(* IEC 61131-3 sources: daoli-st-library/DL_Process (part 41) *)

(* ---- FB_DL_LyoShelfTempRampCtrl.st ---- *)
(*
  Name: FB_DL_LyoShelfTempRampCtrl
  Category: DL_Process
  Version: 1.0.0
  Round: R91 / 2026-11-25
  开源溯源：clean-room 自研（族 制药冻干真空冷冻干燥，ST 开源生态实测 0 命中，无外部代码引入）
  功能：1) 搁板温度斜坡发生器：设定值 fSetpointC 以 fRateUpKmin / fRateDownKmin 的斜率
           逐拍逼近目标温度 fTargetC，每拍增量 = 斜率[K/min] / 60 * fCycleS[s]，
           接近目标时按「不越过目标」截断，天然消除斜坡积分超调。
        2) 超调抑制：实测温度 fActualC 越过目标温度且超出 fOverShootLimitK 并持续 DL_OV_DELAY 后，
           判超调故障并锁码 —— 这是加热回路失控（固态继电器击穿或传感器脱落）的实证判据。
        3) 斜率上下限约束：fRateUpKmin / fRateDownKmin 必须落在 (0.0, DL_RATE_HI_KMIN] 内，
           越域判故障码（斜率为零会让设定值永不到达，斜率过大会撕裂制品冰晶结构）。
  边界条件：1) 非有限值闸：目标温度、实测温度、两路斜率、周期先过 NOT(x > -DL_BIG AND x < DL_BIG)，
           同时拦 NaN 与 Inf；命中即判故障码 0213 并进故障相，
           绝不把 NaN 写进设定值（NaN 一旦进入斜坡状态量会永久污染积分链，R19）。
        2) 周期入参闸（R21）：fCycleS <= 0.0 或非有限时改用缺省 DL_CYCLE_DEF = 0.1 s 并置信息级码 0212，
           不静默改用。
        3) 斜率零闸：两路斜率均须 > DL_EPS，否则判故障码 0214（斜坡永不推进 = 温度控制静默失效）。
        4) 超调判据去抖：超调为瞬时量，必须经 tonOver 去抖后才升级为故障，避免单点尖峰误停。
        5) 单点赋值（R26）：fSetpointC 只在段 7 统一出口写一次；内部设定量 _fSpC 才是逐拍累加的对象。
        6) 故障解除路径：故障相内 xReset 上升沿 AND NOT xFault AND 入参有限 → 清锁存回待机，
           回待机后设定值跟随实测温度重新起步（无扰切换），不从零开始。
        7) 状态机兜底：CASE 全态覆盖 + ELSE 强制回故障相并置码 0217、清全部输出。
  量纲自证：斜率 [K/min] / 60 [s/min] * fCycleS [s] = 每拍增量 [K]，
           与 fSetpointC / fTargetC / fOverShootLimitK 同量纲 [K]（degC 差值以 K 计），量纲合法。
  码表 Error codes（本件子带 0091_021x，故障级一律 3 行内置 _uFault/_bFault/_eState）:
    16#0091_0211 信息级：使能关闭，设定值冻结在当下（不置故障位）
    16#0091_0212 信息级：周期入参非法，已按缺省 0.1 s 折算（不置故障位）
    16#0091_0213 故障级：温度或斜率入参非有限（NaN / Inf）
    16#0091_0214 故障级：斜率组态越域（为零或超物理上限）
    16#0091_0215 故障级：实测温度超调越限（加热回路失控判据）
    16#0091_0216 故障级：外部故障输入 xFault
    16#0091_0217 故障级：状态机落 ELSE 兜底（非法相位 ID）

  修订历史 Revision :
    2026-11-25  v1.0.0  R91 首版
*)

TYPE E_DL_LyoShelfRampState :
(
    eLyoRampIdle  := 0,     // 待机：使能关闭，设定值冻结 / Idle, disabled and setpoint frozen
    eLyoRampHeat  := 10,    // 升温：设定值按升斜率逼近目标 / Heating, setpoint ramps up to target
    eLyoRampCool  := 20,    // 降温：设定值按降斜率逼近目标 / Cooling, setpoint ramps down to target
    eLyoRampHold  := 30,    // 保持：设定值已达目标，进入保温带 / Hold, setpoint on target within the band
    eLyoRampFault := 90     // 故障：锁存待解除 / Fault, latched awaiting release
);
END_TYPE

FUNCTION_BLOCK FB_DL_LyoShelfTempRampCtrl
VAR_INPUT
    xEnable        : BOOL;    // 斜坡控制使能 [bool] / Ramp control enable [bool]
    xReset         : BOOL;    // 故障复位（上升沿有效）[bool] / Fault reset, rising edge [bool]
    xFault         : BOOL;    // 外部故障汇总 [bool] / External fault aggregate [bool]
    fTargetC       : REAL;    // 搁板目标温度 [degC] / Shelf target temperature [degC]
    fActualC       : REAL;    // 搁板实测温度 [degC] / Shelf measured temperature [degC]
    fRateUpKmin    : REAL;    // 允许升温斜率 [K/min] / Permitted heating rate [K/min]
    fRateDownKmin  : REAL;    // 允许降温斜率 [K/min] / Permitted cooling rate [K/min]
    fCycleS        : REAL;    // 任务周期 [s] / Task cycle time [s]
    fBandK         : REAL;    // 到温判定带宽 [K] / At-target band width [K]
    fOverShootLimitK : REAL;  // 允许超调量 [K] / Permitted overshoot [K]
END_VAR
VAR_OUTPUT
    fSetpointC     : REAL;    // 搁板温度设定值 [degC] / Shelf temperature setpoint [degC]
    xHeating       : BOOL;    // 升温方向标志 [bool] / Heating direction flag [bool]
    xCooling       : BOOL;    // 降温方向标志 [bool] / Cooling direction flag [bool]
    xInBand        : BOOL;    // 已进入到温带 [bool] / Within the at-target band [bool]
    xOverShoot     : BOOL;    // 超调越限标志（已去抖）[bool] / Overshoot flag, debounced [bool]
    eState         : E_DL_LyoShelfRampState;   // 状态出口，段尾单点映射 / State outlet, single-point mapped
    nErrId         : UDINT;   // 事件码，0 = 无事件 / Event code, 0 = none
END_VAR
VAR
    tonOver        : TON;     // 超调去抖定时 [TIME] / Overshoot debounce timer
    rtReset        : R_TRIG;  // 复位上升沿检测 [bool] / Reset rising edge detector
    _eState        : E_DL_LyoShelfRampState := E_DL_LyoShelfRampState.eLyoRampIdle;   // 内部相位（CASE 唯一写入目标）
    _fSpC          : REAL := 0.0;   // 内部设定值状态量（逐拍累加对象）[degC] / Internal setpoint state [degC]
    _fStepK        : REAL := 0.0;   // 本拍温度增量 [K] / Temperature increment this cycle [K]
    _fCycleUseS    : REAL := 0.1;   // 实际使用的周期值 [s] / Cycle time actually used [s]
    _bFinOk        : BOOL := FALSE; // 实值入参有限性总闸结果 / Finiteness gate aggregate result
    _bRateOk       : BOOL := FALSE; // 斜率组态域闸结果 / Ramp rate domain gate result
    _bCycleBad     : BOOL := FALSE; // 周期入参非法标志 [bool] / Cycle input invalid flag [bool]
    _bOverRaw      : BOOL := FALSE; // 超调原始判据（未去抖）[bool] / Raw overshoot criterion
    _bFault        : BOOL := FALSE; // 故障锁存位 [bool] / Latched fault flag [bool]
    _bSpInit       : BOOL := FALSE; // 设定值已初始化标志 [bool] / Setpoint initialised flag [bool]
    _uInfo         : UDINT := 16#0000_0000;   // 信息码，每拍重算 / Info code, recomputed every cycle
    _uFault        : UDINT := 16#0000_0000;   // 故障码锁存 / Latched fault code
END_VAR
VAR CONSTANT
    DL_EPS         : REAL := 1.0E-9;      // 数值零闸阈值 [-] / Numeric zero gate threshold [-]
    DL_BIG         : REAL := 1.0E12;      // 非有限值闸量级上限 [-] / Finiteness gate magnitude [-]
    DL_CYCLE_DEF   : REAL := 0.1;         // 缺省任务周期 [s] / Default task cycle time [s]
    DL_CYCLE_MIN   : REAL := 0.001;       // 周期合理下限 [s] / Cycle time reasonable low bound [s]
    DL_CYCLE_MAX   : REAL := 10.0;        // 周期合理上限 [s] / Cycle time reasonable high bound [s]
    DL_SEC_PER_MIN : REAL := 60.0;        // 分钟到秒的时基折算 [s/min] / Seconds per minute [s/min]
    DL_RATE_HI_KMIN: REAL := 10.0;        // 允许斜率物理上限 [K/min] / Ramp rate physical upper bound [K/min]
    DL_OV_DELAY    : TIME := T#10S;       // 超调去抖窗 [TIME] / Overshoot debounce window [TIME]
    DL_T_SPAN      : REAL := 300.0;       // 温度量级闸跨度 [degC] / Temperature magnitude gate span [degC]
END_VAR

(* —— 段 0：单拍量预清零（锁存量 _uFault/_bFault/_bSpInit 不入清单，R187①） —— *)
_uInfo := 16#0000_0000;                     // 信息码每拍重算 / Info code recomputed
nErrId := 16#0000_0000;                     // 事件码缺省无事件 / Event code defaults to none

(* —— 段 1：周期入参闸（R21：非法周期不静默，改用缺省并置信息码） —— *)
_bCycleBad := NOT (fCycleS > -DL_BIG AND fCycleS < DL_BIG)
              OR (fCycleS < DL_CYCLE_MIN) OR (fCycleS > DL_CYCLE_MAX);
IF _bCycleBad THEN
    _fCycleUseS := DL_CYCLE_DEF;            // 非法周期一律用缺省 0.1 s
    _uInfo := 16#0091_0212;                 // 信息级：周期入参非法，已用缺省（不置故障位）
ELSE
    _fCycleUseS := fCycleS;                 // 合法周期原值使用
END_IF

(* —— 段 2：非有限值闸与斜率域闸（R19：不把 NaN 写进斜坡状态量） —— *)
_bFinOk := (fTargetC > -DL_BIG) AND (fTargetC < DL_BIG)
           AND (fActualC > -DL_BIG) AND (fActualC < DL_BIG)
           AND (fRateUpKmin > -DL_BIG) AND (fRateUpKmin < DL_BIG)
           AND (fRateDownKmin > -DL_BIG) AND (fRateDownKmin < DL_BIG)
           AND (fBandK > -DL_BIG) AND (fBandK < DL_BIG)
           AND (fOverShootLimitK > -DL_BIG) AND (fOverShootLimitK < DL_BIG);
_bRateOk := (fRateUpKmin > DL_EPS) AND (fRateUpKmin <= DL_RATE_HI_KMIN)
            AND (fRateDownKmin > DL_EPS) AND (fRateDownKmin <= DL_RATE_HI_KMIN)
            AND (fBandK > DL_EPS) AND (fOverShootLimitK > DL_EPS)
            AND (ABS(fTargetC) <= DL_T_SPAN) AND (ABS(fActualC) <= DL_T_SPAN);

(* —— 段 3：超调原始判据（仅升温方向有意义：实测高于目标且超出允许量） —— *)
_bOverRaw := _bFinOk AND _bRateOk
             AND ((fActualC - fTargetC) > fOverShootLimitK);

(* —— 段 4：边沿与定时器无条件周期刷新（R7：调用语句不得置于 IF/CASE 内） —— *)
rtReset(CLK := xReset);                                             // 复位上升沿，每拍必调
tonOver(IN := _bOverRaw AND (NOT _bFault), PT := DL_OV_DELAY);      // 超调去抖

(* —— 段 5：全局故障拦截（优先级最高；已锁存则不再改写码值，禁同拍抹除） —— *)
IF xFault AND (NOT _bFault) THEN
    _uFault := 16#0091_0216;                // 故障级：外部故障输入
    _bFault := TRUE;                        // 锁存（3 行内置，R45 配对）
    _eState := E_DL_LyoShelfRampState.eLyoRampFault;
END_IF
IF (NOT _bFinOk) AND (NOT _bFault) THEN
    _uFault := 16#0091_0213;                // 故障级：入参非有限（独立成因，R190）
    _bFault := TRUE;                        // 锁存
    _eState := E_DL_LyoShelfRampState.eLyoRampFault;
END_IF
IF (NOT _bRateOk) AND _bFinOk AND (NOT _bFault) THEN
    _uFault := 16#0091_0214;                // 故障级：斜率组态越域（独立成因，R190）
    _bFault := TRUE;                        // 锁存
    _eState := E_DL_LyoShelfRampState.eLyoRampFault;
END_IF
IF tonOver.Q AND (NOT _bFault) THEN
    _uFault := 16#0091_0215;                // 故障级：实测温度超调越限
    _bFault := TRUE;                        // 锁存
    _eState := E_DL_LyoShelfRampState.eLyoRampFault;
END_IF

(* —— 段 6：设定值起步（首次使能或无扰复位时以实测温度初始化，避免设定值从零跳变） —— *)
IF (NOT _bSpInit) AND _bFinOk THEN
    _fSpC := fActualC;                      // 无扰起步：设定值跟随实测温度
    _bSpInit := TRUE;                       // 标记已初始化
END_IF

(* —— 段 7：相位机（只做迁移与内部设定值更新；出口在段 9 单点映射） —— *)
CASE _eState OF

E_DL_LyoShelfRampState.eLyoRampIdle:
    IF NOT xEnable THEN
        _uInfo := 16#0091_0211;             // 信息级：使能关闭，设定值冻结（不置故障位）
    ELSIF (fTargetC - _fSpC) > fBandK THEN
        _eState := E_DL_LyoShelfRampState.eLyoRampHeat;       // 目标高于设定值：进升温相
    ELSIF (_fSpC - fTargetC) > fBandK THEN
        _eState := E_DL_LyoShelfRampState.eLyoRampCool;       // 目标低于设定值：进降温相
    ELSE
        _eState := E_DL_LyoShelfRampState.eLyoRampHold;       // 已在带内：进保持相
    END_IF

E_DL_LyoShelfRampState.eLyoRampHeat:
    IF (NOT xEnable) OR _bFault THEN
        _uInfo := 16#0091_0211;             // 信息级：失能即冻结设定值
        _eState := E_DL_LyoShelfRampState.eLyoRampIdle;
    ELSE
        _fStepK := fRateUpKmin / DL_SEC_PER_MIN * _fCycleUseS;                 // 每拍升温增量 [K]
        _fSpC := _fSpC + _fStepK;                                             // 累加
        IF _fSpC >= fTargetC THEN
            _fSpC := fTargetC;              // 不越过目标：天然消除斜坡超调
            _eState := E_DL_LyoShelfRampState.eLyoRampHold;
        END_IF
    END_IF

E_DL_LyoShelfRampState.eLyoRampCool:
    IF (NOT xEnable) OR _bFault THEN
        _uInfo := 16#0091_0211;             // 信息级：失能即冻结设定值
        _eState := E_DL_LyoShelfRampState.eLyoRampIdle;
    ELSE
        _fStepK := fRateDownKmin / DL_SEC_PER_MIN * _fCycleUseS;               // 每拍降温增量 [K]
        _fSpC := _fSpC - _fStepK;                                             // 累减
        IF _fSpC <= fTargetC THEN
            _fSpC := fTargetC;              // 不越过目标：天然消除斜坡超调
            _eState := E_DL_LyoShelfRampState.eLyoRampHold;
        END_IF
    END_IF

E_DL_LyoShelfRampState.eLyoRampHold:
    IF (NOT xEnable) OR _bFault THEN
        _uInfo := 16#0091_0211;             // 信息级：失能即回待机
        _eState := E_DL_LyoShelfRampState.eLyoRampIdle;
    ELSIF (fTargetC - _fSpC) > fBandK THEN
        _eState := E_DL_LyoShelfRampState.eLyoRampHeat;       // 目标抬高：重返升温相（判据在钉住之前取）
    ELSIF (_fSpC - fTargetC) > fBandK THEN
        _eState := E_DL_LyoShelfRampState.eLyoRampCool;       // 目标压低：重返降温相（判据在钉住之前取）
    ELSE
        _fSpC := fTargetC;                  // 带内才钉住设定值（避免判据恒真）
    END_IF

E_DL_LyoShelfRampState.eLyoRampFault:
    IF rtReset.Q AND (NOT xFault) AND _bFinOk AND _bRateOk THEN
        _bFault := FALSE;                   // 解除路径：复位沿 + 外部故障消失 + 入参与组态合法（可达，R188）
        _uFault := 16#0000_0000;            // 清锁存码
        _bSpInit := FALSE;                  // 强制无扰重启：设定值重新跟随实测温度
        _eState := E_DL_LyoShelfRampState.eLyoRampIdle;       // 回待机
    END_IF

ELSE
    _uFault := 16#0091_0217;                // 故障级：非法相位 ID 兜底
    _bFault := TRUE;                        // 锁存
    _eState := E_DL_LyoShelfRampState.eLyoRampFault;          // 强制回故障相

END_CASE

(* —— 段 8：后置段（设定值域兜底：非有限或越量级一律回落到实测温度） —— *)
IF NOT (_fSpC > -DL_BIG AND _fSpC < DL_BIG) THEN
    _fSpC := fActualC;                      // 内部状态自检：非有限即回落实测值
END_IF
(* —— 段 8.5：出口值域二阶终闸（R19 二阶形态）——
   一次闸的回退源是 fActualC，而 fActualC 本身也可能是非有限值（入参 NaN/Inf），
   回退后仍为 NaN，且 ABS(NaN) > DL_T_SPAN 恒假会绕过越量级钳制，NaN 直穿设定值出口。
   故必须对「回退之后」的值再做一次判据与钳制，才真正闸断实值通路。 *)
IF NOT (_fSpC >= -DL_T_SPAN AND _fSpC <= DL_T_SPAN) THEN
    _fSpC := 0.0;                           // 双源皆非有限：0 degC 安全位 / Both sources non-finite: 0 degC safe
END_IF
IF ABS(_fSpC) > DL_T_SPAN THEN
    _fSpC := LIMIT(-DL_T_SPAN, _fSpC, DL_T_SPAN);   // 越量级钳制，防积分链发散
END_IF

(* —— 段 9：出口单点映射（名实同源；方向位由设定值与目标差导出，故障侧全清） —— *)
IF _bFault THEN
    IF (fActualC >= -DL_T_SPAN) AND (fActualC <= DL_T_SPAN) THEN
        fSetpointC := fActualC;             // 故障侧优先回落实测温度（有限时保持原语义：冻结在实测）
    ELSE
        fSetpointC := _fSpC;                // 实测非有限时回落到已过二阶终闸的安全值，绝不输出 NaN
    END_IF;
    xHeating := FALSE;                      // 故障侧方向位清零
    xCooling := FALSE;                      // 故障侧方向位清零
    xInBand := FALSE;                       // 故障侧到温位清零
ELSE
    fSetpointC := _fSpC;                    // 正常侧设定值出口
    xHeating := (_eState = E_DL_LyoShelfRampState.eLyoRampHeat);      // 升温方向位
    xCooling := (_eState = E_DL_LyoShelfRampState.eLyoRampCool);      // 降温方向位
    xInBand := (_eState = E_DL_LyoShelfRampState.eLyoRampHold)        // 到温带：保持相且实测在带内
               AND (ABS(fActualC - fTargetC) <= fBandK);
END_IF
xOverShoot := tonOver.Q;                    // 超调位出口（已去抖）
eState := _eState;                          // 状态出口单点映射
IF _bFault THEN
    nErrId := _uFault;                      // 故障锁存码回放（不在故障相按当下输入重推断）
ELSE
    nErrId := _uInfo;                       // 信息码
END_IF

END_FUNCTION_BLOCK

(* ---- FB_DL_LyoVacuumPullSeq.st ---- *)
(*
  Name: FB_DL_LyoVacuumPullSeq
  Category: DL_Process
  Version: 1.0.0
  Round: R91 / 2026-11-25
  开源溯源：clean-room 自研（族 制药冻干真空冷冻干燥，ST 开源生态实测 0 命中，无外部代码引入）
  功能：1) 抽真空状态机，六相推进：待机 → 粗抽 → 精抽 → 保持 → 就绪 → （通气）。
           待机相等 xStart 上升沿；腔体压力已低于粗抽目标时跳过粗抽相（信息级码 0231 声明跳过）；
           粗抽相开粗抽泵阀组，压力降到 fRoughTargetMbar 即转精抽；精抽相关粗抽阀、开精抽阀，
           压力降到 fFineTargetMbar 即转保持相；保持相关全部抽气、观察 tHoldS 内压力升幅，
           升幅 <= fHoldRiseMaxMbar 判真空保持合格，置 xHoldOk 并进就绪相；
           就绪相保持 xReady 直到 xStart 撤下；撤令后进通气相复压并回待机。
        2) 泵故障兜底：粗抽/精抽/保持三相内，泵运行反馈丢失或泵过载上升即锁码 0237 并立即进故障相，
           同时撤销全部抽气命令、不打开通气阀（避免带故障强行复压把油雾带入腔体）。
        3) 每相独立超时 + 整序总超时：四个相定时器各配一个「定时 + 裕量」超时点，
           tonTotal 兜底整序总时长；保持相另配真空上升超限判据（0234）与稳定超时（0235）双归因。
  边界条件：1) 非有限值闸：压力、三个目标限值先过 NOT(x > -DL_BIG AND x < DL_BIG)，同时拦 NaN 与 Inf；
           命中即锁码 0239 进故障相，绝不把 NaN 拿去与真空目标比较（NaN 比较恒假会让抽气永不停止，R19）。
        2) 组态域闸：三个压力阈须满足 0.0 < fFineTargetMbar < fRoughTargetMbar（真空度方向由粗到精），
           fHoldRiseMaxMbar > DL_EPS，越域锁码 0239（组态错误与入参非有限共用同一归因码前缀，
           但内部用两个独立成员区分，见 _bCfgOk / _bFinOk）。
        3) 压力单调性：抽气相内压力不得上升；若在粗抽/精抽相检测到压力高于本相入口压力且超过
           DL_PRESS_TOL，视为泵失效实测证据，锁码 0232 / 0233（与超时归因区分：这里不是等不到，而是反向）。
        4) 时间参数零闸：tRoughS / tFineS / tHoldS <= T#0S 时对应相定时器立即置 Q（等价跳过），
           属调试合法组态；但保持相零窗会使升幅判据恒成立，故保持相入口对 tHoldS 做显式零闸 → 锁码 0235。
        5) 定时器周期刷新（R7）：八个 TON 与复位边沿全部在 CASE 之外无条件调用。
        6) 故障解除路径：故障相内 xReset 上升沿 AND NOT xFault AND 入参/组态合法 → 清锁存回待机，
           回待机后必须重新给 xStart 上升沿才能再启动（不自恢复）。
        7) 状态机兜底：CASE 全态覆盖 + ELSE 强制回故障相并置码 0240、清全部输出。
        8) 输出安全初值（R25）：三个阀门命令初值 FALSE、xReady 初值 FALSE，待机相显式赋值。
  量纲自证：fChamberPressMbar / fRoughTargetMbar / fFineTargetMbar / fHoldRiseMaxMbar 全为压力 [mbar]，
           比较两侧同量纲；升幅 = 保持末压力 − 保持初压力，仍为 [mbar]；
           所有时间引脚为 [TIME]，相超时点 = [TIME] + [TIME] = [TIME]，与 TON 的 PT 同量纲。
  码表 Error codes（本件子带 0091_024x，故障级一律 3 行内置 _uFault/_bFault/_eState）:
    16#0091_0231 信息级：腔体压力已低于粗抽目标，跳过粗抽相（不置故障位）
    16#0091_0232 故障级：粗抽相超时（定时到但未达粗抽目标）
    16#0091_0233 故障级：精抽相超时（定时到但未达精抽目标）
    16#0091_0234 故障级：保持相真空度上升超限（泄漏或放气）
    16#0091_0235 故障级：保持相超时或保持窗为零（压力未稳定/判据恒真）
    16#0091_0236 故障级：整序总超时
    16#0091_0237 故障级：泵运行反馈丢失或泵过载
    16#0091_0238 故障级：外部故障输入 xFault
    16#0091_0239 故障级：压力/限值入参非有限，或压力阈组态越域
    16#0091_0240 故障级：状态机落 ELSE 兜底（非法相位 ID）
    16#0091_0241 信息级：就绪保持中，等待撤令（不置故障位）
    16#0091_0242 信息级：通气复压相进行中（不置故障位）
    16#0091_0243 信息级：泵未就绪（无运行反馈或过载），暂不启动抽气（不置故障位）
    16#0091_0244 故障级：粗抽相压力反向上升（泵失效实证，与超时成因分离）
    16#0091_0245 故障级：精抽相压力反向上升（泄漏或阀未开，与超时成因分离）
    16#0091_0246 故障级：通气相超时（复压未完成）

  修订历史 Revision :
    2026-11-25  v1.0.0  R91 首版
*)

TYPE E_DL_LyoVacuumPullState :
(
    eLyoVacIdle  := 0,      // 待机：等启动上升沿 / Idle, awaiting the start rising edge
    eLyoVacRough := 10,     // 粗抽：粗抽泵组开，降到粗抽目标 / Rough pull, pump group on
    eLyoVacFine  := 20,     // 精抽：关粗抽阀开精抽阀，降到精抽目标 / Fine pull, fine valve open
    eLyoVacHold  := 30,     // 保持：关全部抽气，测压力升幅 / Hold, all pumping off, rise measured
    eLyoVacReady := 40,     // 就绪：真空保持合格，保持到位 / Ready, vacuum hold accepted
    eLyoVacVent  := 50,     // 通气：开通气阀复压回待机 / Vent, repressurising back to idle
    eLyoVacFault := 90      // 故障：锁存待解除 / Fault, latched awaiting release
);
END_TYPE

FUNCTION_BLOCK FB_DL_LyoVacuumPullSeq
VAR_INPUT
    xStart           : BOOL;   // 抽真空启动指令（上升沿有效）[bool] / Vacuum pull start, edge triggered [bool]
    xReset           : BOOL;   // 故障复位（上升沿有效）[bool] / Fault reset, rising edge [bool]
    xFault           : BOOL;   // 外部故障汇总 [bool] / External fault aggregate [bool]
    xPumpRunFb       : BOOL;   // 真空泵运行反馈 [bool] / Vacuum pump running feedback [bool]
    xPumpOverload    : BOOL;   // 真空泵过载信号 [bool] / Vacuum pump overload signal [bool]
    fChamberPressMbar : REAL;  // 腔体实测压力 [mbar] / Measured chamber pressure [mbar]
    fRoughTargetMbar : REAL;   // 粗抽目标压力 [mbar] / Rough pull target pressure [mbar]
    fFineTargetMbar  : REAL;   // 精抽目标压力 [mbar] / Fine pull target pressure [mbar]
    fHoldRiseMaxMbar : REAL;   // 保持相允许压力升幅 [mbar] / Permitted pressure rise during hold [mbar]
    tRoughS          : TIME;   // 粗抽相设定时长 [TIME] / Rough pull phase duration [TIME]
    tFineS           : TIME;   // 精抽相设定时长 [TIME] / Fine pull phase duration [TIME]
    tHoldS           : TIME;   // 保持相设定时长 [TIME] / Hold phase duration [TIME]
END_VAR
VAR_OUTPUT
    xRoughValveCmd   : BOOL;   // 粗抽阀命令（安全侧：故障时关）[bool] / Rough valve command, fail-safe [bool]
    xFineValveCmd    : BOOL;   // 精抽阀命令（安全侧：故障时关）[bool] / Fine valve command, fail-safe [bool]
    xVentValveCmd    : BOOL;   // 通气阀命令（安全侧：故障时关）[bool] / Vent valve command, fail-safe [bool]
    xHoldOk          : BOOL;   // 真空保持判据通过（跨相保持）[bool] / Vacuum hold accepted, held across phases [bool]
    xReady           : BOOL;   // 抽真空就绪保持位 [bool] / Vacuum ready held flag [bool]
    xBusy            : BOOL;   // 抽真空进行中 [bool] / Vacuum pull busy [bool]
    eState           : E_DL_LyoVacuumPullState;   // 状态出口，段尾单点映射 / State outlet, single-point mapped
    nErrId           : UDINT;  // 事件码，0 = 无事件 / Event code, 0 = none
END_VAR
VAR
    tonRough         : TON;    // 粗抽相正常定时 [TIME] / Rough pull phase timer
    tonRoughOv       : TON;    // 粗抽相超时定时 [TIME] / Rough pull phase overrun timer
    tonFine          : TON;    // 精抽相正常定时 [TIME] / Fine pull phase timer
    tonFineOv        : TON;    // 精抽相超时定时 [TIME] / Fine pull phase overrun timer
    tonHold          : TON;    // 保持相正常定时 [TIME] / Hold phase timer
    tonHoldOv        : TON;    // 保持相超时定时 [TIME] / Hold phase overrun timer
    tonVent          : TON;    // 通气相正常定时 [TIME] / Vent phase timer
    tonVentOv        : TON;    // 通气相超时定时 [TIME] / Vent phase overrun timer
    tonTotal         : TON;    // 整序总超时定时 [TIME] / Whole-sequence total timeout timer
    rtStart          : R_TRIG; // 启动上升沿检测 [bool] / Start rising edge detector
    rtReset          : R_TRIG; // 复位上升沿检测 [bool] / Reset rising edge detector
    _eState          : E_DL_LyoVacuumPullState := E_DL_LyoVacuumPullState.eLyoVacIdle;   // 内部相位（CASE 唯一写入目标）
    _fPressEntryMbar : REAL := 0.0;   // 本相入口压力快照 [mbar] / Pressure snapshot at phase entry [mbar]
    _fHoldStartMbar  : REAL := 0.0;   // 保持相起点压力快照 [mbar] / Pressure snapshot at hold start [mbar]
    _fRiseMbar       : REAL := 0.0;   // 保持相压力升幅 [mbar] / Pressure rise during the hold phase [mbar]
    _bFinOk          : BOOL := FALSE; // 实值入参有限性总闸结果 / Finiteness gate aggregate result
    _bCfgOk          : BOOL := FALSE; // 压力阈组态域闸结果 / Pressure threshold domain gate result
    _bPumpOk         : BOOL := FALSE; // 泵健康（运行反馈有且无过载）[bool] / Pump healthy flag [bool]
    _bActive         : BOOL := FALSE; // 序激活（粗抽至通气五相之一）[bool] / Sequence active flag [bool]
    _bHoldL          : BOOL := FALSE; // 保持合格位锁存（跨相保持）[bool] / Hold-accepted latch [bool]
    _bFault          : BOOL := FALSE; // 故障锁存位 [bool] / Latched fault flag [bool]
    _uInfo           : UDINT := 16#0000_0000;   // 信息码，每拍重算 / Info code, recomputed every cycle
    _uFault          : UDINT := 16#0000_0000;   // 故障码锁存 / Latched fault code
END_VAR
VAR CONSTANT
    DL_EPS         : REAL := 1.0E-9;      // 数值零闸阈值 [-] / Numeric zero gate threshold [-]
    DL_BIG         : REAL := 1.0E12;      // 非有限值闸量级上限 [-] / Finiteness gate magnitude [-]
    DL_PRESS_TOL   : REAL := 0.05;        // 抽气相压力反向容差 [mbar] / Reverse-trend tolerance while pumping [mbar]
    DL_P_HI        : REAL := 1100.0;      // 压力量级闸上限（略高于常压）[mbar] / Pressure magnitude gate upper bound [mbar]
    DL_OVER_MARGIN : TIME := T#60S;       // 相超时相对正常定时的裕量 [TIME] / Phase overrun margin [TIME]
    DL_TOTAL_MAX   : TIME := T#4H;        // 整序总超时上限 [TIME] / Whole-sequence total timeout [TIME]
    DL_ZERO_PRES   : REAL := 0.0;         // 压力零基准 [mbar] / Zero pressure reference [mbar]
END_VAR

(* —— 段 0：单拍量预清零（锁存量 _uFault/_bFault/_bHoldL 不入清单，R187①） —— *)
_uInfo := 16#0000_0000;                     // 信息码每拍重算 / Info code recomputed
nErrId := 16#0000_0000;                     // 事件码缺省无事件 / Event code defaults to none

(* —— 段 1：非有限值闸与组态域闸（R19：不拿 NaN 去比较真空目标） —— *)
_bFinOk := (fChamberPressMbar > -DL_BIG) AND (fChamberPressMbar < DL_BIG)
           AND (fRoughTargetMbar > -DL_BIG) AND (fRoughTargetMbar < DL_BIG)
           AND (fFineTargetMbar > -DL_BIG) AND (fFineTargetMbar < DL_BIG)
           AND (fHoldRiseMaxMbar > -DL_BIG) AND (fHoldRiseMaxMbar < DL_BIG);
_bCfgOk := (fFineTargetMbar > DL_EPS)                       // 精抽目标须为正压
           AND (fFineTargetMbar < fRoughTargetMbar)         // 精抽必须比粗抽更深（方向由粗到精）
           AND (fRoughTargetMbar < DL_P_HI)                 // 粗抽目标须在压力量级内
           AND (fHoldRiseMaxMbar > DL_EPS);                 // 允许升幅须组态为正

(* —— 段 2：泵健康判据（运行反馈 + 过载；过载优先） —— *)
_bPumpOk := xPumpRunFb AND (NOT xPumpOverload);

(* —— 段 3：派生态（序激活、保持升幅） —— *)
_bActive := (_eState = E_DL_LyoVacuumPullState.eLyoVacRough)
            OR (_eState = E_DL_LyoVacuumPullState.eLyoVacFine)
            OR (_eState = E_DL_LyoVacuumPullState.eLyoVacHold)
            OR (_eState = E_DL_LyoVacuumPullState.eLyoVacReady)
            OR (_eState = E_DL_LyoVacuumPullState.eLyoVacVent);
_fRiseMbar := fChamberPressMbar - _fHoldStartMbar;          // 保持相压力升幅 [mbar]

(* —— 段 4：定时器与边沿无条件周期刷新（R7：调用语句不得置于 IF/CASE 内） —— *)
rtStart(CLK := xStart);                                                                   // 启动上升沿，每拍必调
rtReset(CLK := xReset);                                                                   // 复位上升沿，每拍必调
tonRough(IN := (_eState = E_DL_LyoVacuumPullState.eLyoVacRough), PT := tRoughS);          // 粗抽相正常定时
tonRoughOv(IN := (_eState = E_DL_LyoVacuumPullState.eLyoVacRough),
           PT := tRoughS + DL_OVER_MARGIN);                                               // 粗抽相超时点
tonFine(IN := (_eState = E_DL_LyoVacuumPullState.eLyoVacFine), PT := tFineS);             // 精抽相正常定时
tonFineOv(IN := (_eState = E_DL_LyoVacuumPullState.eLyoVacFine),
          PT := tFineS + DL_OVER_MARGIN);                                                 // 精抽相超时点
tonHold(IN := (_eState = E_DL_LyoVacuumPullState.eLyoVacHold), PT := tHoldS);             // 保持相正常定时
tonHoldOv(IN := (_eState = E_DL_LyoVacuumPullState.eLyoVacHold),
          PT := tHoldS + DL_OVER_MARGIN);                                                 // 保持相超时点
tonVent(IN := (_eState = E_DL_LyoVacuumPullState.eLyoVacVent), PT := tRoughS);            // 通气相正常定时（借用粗抽时长作复压窗）
tonVentOv(IN := (_eState = E_DL_LyoVacuumPullState.eLyoVacVent),
          PT := tRoughS + DL_OVER_MARGIN);                                                // 通气相超时点
tonTotal(IN := _bActive, PT := DL_TOTAL_MAX);                                             // 整序总超时

(* —— 段 5：全局故障拦截（优先级最高；已锁存则不再改写码值，禁同拍抹除） —— *)
IF xFault AND (NOT _bFault) THEN
    _uFault := 16#0091_0238;                // 故障级：外部故障输入
    _bFault := TRUE;                        // 锁存（3 行内置，R45 配对）
    _eState := E_DL_LyoVacuumPullState.eLyoVacFault;
END_IF
IF ((NOT _bFinOk) OR (NOT _bCfgOk)) AND (NOT _bFault) THEN
    _uFault := 16#0091_0239;                // 故障级：入参非有限或压力阈组态越域（同一码，成员已分离）
    _bFault := TRUE;                        // 锁存
    _eState := E_DL_LyoVacuumPullState.eLyoVacFault;
END_IF
IF tonTotal.Q AND _bActive AND (NOT _bFault) THEN
    _uFault := 16#0091_0236;                // 故障级：整序总超时
    _bFault := TRUE;                        // 锁存
    _eState := E_DL_LyoVacuumPullState.eLyoVacFault;
END_IF
IF (NOT _bPumpOk) AND _bActive AND (NOT _bFault)
   AND (_eState <> E_DL_LyoVacuumPullState.eLyoVacVent) THEN
    _uFault := 16#0091_0237;                // 故障级：泵反馈丢失或过载（通气相不需泵，故排除）
    _bFault := TRUE;                        // 锁存
    _eState := E_DL_LyoVacuumPullState.eLyoVacFault;
END_IF

(* —— 段 6：相位机（只做迁移与锁存；出口在段 8 单点映射） —— *)
CASE _eState OF

E_DL_LyoVacuumPullState.eLyoVacIdle:
    IF NOT xStart THEN
        _bHoldL := FALSE;                   // 撤令即清保持合格位，为下次抽真空重新武装
        _fPressEntryMbar := fChamberPressMbar;   // 待机相刷新入口压力快照（有限性由段 5 保证）
    ELSIF rtStart.Q AND _bFinOk AND _bCfgOk THEN
        _bHoldL := FALSE;                   // 新序开始：清保持合格位
        _fPressEntryMbar := fChamberPressMbar;   // 捕获入口压力，供粗抽反向判据使用
        IF fChamberPressMbar <= fRoughTargetMbar THEN
            _uInfo := 16#0091_0231;         // 信息级：已低于粗抽目标，声明跳过粗抽相
            _eState := E_DL_LyoVacuumPullState.eLyoVacFine;      // 直接进精抽相
        ELSE
            _eState := E_DL_LyoVacuumPullState.eLyoVacRough;     // 进粗抽相
        END_IF
    ELSIF NOT _bPumpOk THEN
        _uInfo := 16#0091_0243;             // 信息级：泵未就绪，暂不启动（不置故障位）
    END_IF

E_DL_LyoVacuumPullState.eLyoVacRough:
    IF tonRoughOv.Q THEN
        _uFault := 16#0091_0232;            // 故障级：粗抽相超时
        _bFault := TRUE;                    // 锁存
        _eState := E_DL_LyoVacuumPullState.eLyoVacFault;
    ELSIF (fChamberPressMbar - _fPressEntryMbar) > DL_PRESS_TOL THEN
        _uFault := 16#0091_0244;            // 故障级：粗抽中压力反向上升（泵失效实证，独立成因）
        _bFault := TRUE;                    // 锁存
        _eState := E_DL_LyoVacuumPullState.eLyoVacFault;
    ELSIF fChamberPressMbar <= fRoughTargetMbar THEN
        _fPressEntryMbar := fChamberPressMbar;                   // 达粗抽目标：刷新入口快照（迁移前一次性）
        _eState := E_DL_LyoVacuumPullState.eLyoVacFine;          // 进精抽相
    END_IF

E_DL_LyoVacuumPullState.eLyoVacFine:
    IF tonFineOv.Q THEN
        _uFault := 16#0091_0233;            // 故障级：精抽相超时
        _bFault := TRUE;                    // 锁存
        _eState := E_DL_LyoVacuumPullState.eLyoVacFault;
    ELSIF (fChamberPressMbar - _fPressEntryMbar) > DL_PRESS_TOL THEN
        _uFault := 16#0091_0245;            // 故障级：精抽中压力反向上升（泄漏或阀未开，独立成因）
        _bFault := TRUE;                    // 锁存
        _eState := E_DL_LyoVacuumPullState.eLyoVacFault;
    ELSIF fChamberPressMbar <= fFineTargetMbar THEN
        _fHoldStartMbar := fChamberPressMbar;                    // 达精抽目标：捕获保持相起点压力
        _eState := E_DL_LyoVacuumPullState.eLyoVacHold;          // 进保持相
    END_IF

E_DL_LyoVacuumPullState.eLyoVacHold:
    IF tHoldS <= T#0S THEN
        _uFault := 16#0091_0235;            // 故障级：保持窗为零，升幅判据恒成立（不可接受组态）
        _bFault := TRUE;                    // 锁存
        _eState := E_DL_LyoVacuumPullState.eLyoVacFault;
    ELSIF tonHoldOv.Q THEN
        _uFault := 16#0091_0235;            // 故障级：保持相超时（压力未稳定）
        _bFault := TRUE;                    // 锁存
        _eState := E_DL_LyoVacuumPullState.eLyoVacFault;
    ELSIF tonHold.Q THEN
        IF _fRiseMbar > fHoldRiseMaxMbar THEN
            _uFault := 16#0091_0234;        // 故障级：保持相真空度上升超限（泄漏/放气）
            _bFault := TRUE;                // 锁存
            _eState := E_DL_LyoVacuumPullState.eLyoVacFault;
        ELSE
            _bHoldL := TRUE;                // 真空保持合格：锁存（跨相保持）
            _eState := E_DL_LyoVacuumPullState.eLyoVacReady;     // 进就绪相
        END_IF
    END_IF

E_DL_LyoVacuumPullState.eLyoVacReady:
    IF NOT xStart THEN
        _bHoldL := FALSE;                   // 撤令：清保持合格位并进通气相
        _eState := E_DL_LyoVacuumPullState.eLyoVacVent;
    ELSE
        _uInfo := 16#0091_0241;             // 信息级：就绪保持中，等撤令（不置故障位）
    END_IF

E_DL_LyoVacuumPullState.eLyoVacVent:
    IF tonVentOv.Q THEN
        _uFault := 16#0091_0246;            // 故障级：通气相超时（复压未完成，独立成因）
        _bFault := TRUE;                    // 锁存
        _eState := E_DL_LyoVacuumPullState.eLyoVacFault;
    ELSIF tonVent.Q THEN
        _eState := E_DL_LyoVacuumPullState.eLyoVacIdle;          // 复压完成：回待机
    ELSE
        _uInfo := 16#0091_0242;             // 信息级：通气复压进行中（不置故障位）
    END_IF

E_DL_LyoVacuumPullState.eLyoVacFault:
    IF rtReset.Q AND (NOT xFault) AND _bFinOk AND _bCfgOk THEN
        _bFault := FALSE;                   // 解除路径：复位沿 + 外部故障消失 + 入参/组态合法（可达，R188）
        _uFault := 16#0000_0000;            // 清锁存码
        _bHoldL := FALSE;                   // 保持合格位一并清，避免故障后误报就绪
        _eState := E_DL_LyoVacuumPullState.eLyoVacIdle;          // 回待机，需新上升沿才可再启动
    END_IF

ELSE
    _uFault := 16#0091_0240;                // 故障级：非法相位 ID 兜底
    _bFault := TRUE;                        // 锁存
    _eState := E_DL_LyoVacuumPullState.eLyoVacFault;             // 强制回故障相

END_CASE

(* —— 段 7：后置段（压力快照域兜底：非有限即清零，防污染下拍反向判据） —— *)
IF NOT (_fPressEntryMbar > -DL_BIG AND _fPressEntryMbar < DL_BIG) THEN
    _fPressEntryMbar := DL_ZERO_PRES;       // 内部状态自检：非有限即清零
END_IF
IF NOT (_fHoldStartMbar > -DL_BIG AND _fHoldStartMbar < DL_BIG) THEN
    _fHoldStartMbar := DL_ZERO_PRES;        // 内部状态自检：非有限即清零
END_IF

(* —— 段 8：出口单点映射（名实同源；阀门由状态导出，故障侧一律关阀） —— *)
xRoughValveCmd := (_eState = E_DL_LyoVacuumPullState.eLyoVacRough) AND (NOT _bFault);    // 粗抽阀：仅粗抽相
xFineValveCmd := (_eState = E_DL_LyoVacuumPullState.eLyoVacFine) AND (NOT _bFault);      // 精抽阀：仅精抽相
xVentValveCmd := (_eState = E_DL_LyoVacuumPullState.eLyoVacVent) AND (NOT _bFault);      // 通气阀：仅通气相
xHoldOk := _bHoldL AND (NOT _bFault);                                                    // 保持合格位出口
xReady := (_eState = E_DL_LyoVacuumPullState.eLyoVacReady) AND _bHoldL AND (NOT _bFault);   // 就绪位出口
xBusy := _bActive AND (NOT _bFault);                                                     // 进行中出口
eState := _eState;                                                                       // 状态出口单点映射
IF _bFault THEN
    nErrId := _uFault;                      // 故障锁存码回放（不在故障相按当下输入重推断）
ELSE
    nErrId := _uInfo;                       // 信息码
END_IF

END_FUNCTION_BLOCK

(* ---- FB_DL_MachineGuardAudit.st ---- *)
(*==============================================================================
 * 组件名称 (Component)  : FB_DL_MachineGuardAudit
 * 所属子库 (Sublibrary) : DL_Process
 * 当前版本 (Version)    : 1.0.0
 * 兼容性 (Platform)     : CODESYS 3.5 / TwinCAT 3 / 汇川 InoProShop / Machine Expert
 *                         仅依赖纯 IEC 61131-3 标准元素，零厂商方言
 * 功能描述 (Function)   : 防护门开启审计与批次锁定：门开上升沿 → 若批次活动中
 *                         则按 Holding 语义锁批次并记审计（计数饱和、操作员留痕）→
 *                         Held；恢复需「门已关 + 人工确认」→ RESUMING 核实 →
 *                         NORMAL。开门超 tMaxOpen → VIOLATION 锁存，需操作员标识
 *                         与复位双条件方可解锁。本件只借用 Holding/Held 语义组织
 *                         状态，不属主、不替代整机 PackML 状态机。
 * 溯源 (Origin)         : 道莅 clean-room 防御性实现
 * 本文件内含 (Contains) : TYPE E_DL_GuardAuditState / TYPE E_DL_GuardErr /
 *                         FUNCTION_BLOCK FB_DL_MachineGuardAudit
 * 依赖 (Depends)        : 无 DL_ 内部依赖；Standard.library TON/R_TRIG 实例
 * 红线自检 (Redline)    : 无外部全局变量、无硬件地址直引 ｜ 全变量中英双语同行注释
 *                         计数饱和保护 + 门信号保守处置 ｜ 枚举成员全部显式赋值 ｜
 *                         TON/R_TRIG 每周期无条件调用（仅输入条件化）｜
 *                         CASE 含 ELSE 兜底（ELSE → VIOLATION 锁存 + 锁批次）｜
 *                         禁用系统时间函数（审计时间戳由调用方另行记录）
 * 错误码表 (Codes)      : 16#0005_042B NORMAL
 *                         16#0005_042C HOLDING（批次已锁）
 *                         16#0005_042D HELD（等待恢复确认）
 *                         16#0005_042E VIOLATION（超时锁存，需权限复位）
 *                         16#0005_042F RESUMING（恢复核实）
 * 修订历史 (Revision)   : 2026-11-17  v1.0.0  首版入库 · R27 · 阶段三批 4
 * 验收向量 (Acceptance) : 批次活动中门开 → HOLDING(042C) + bLockBatch → HELD(042D)；
 *                         门关 + bManualConfirm → RESUMING(042F) → NORMAL(042B)；
 *                         开门超 tMaxOpen → VIOLATION(042E)，空 sOperId 复位无效
 *============================================================================*)

(*-----------------------------------------------------------------------------
 * 枚举: E_DL_GuardAuditState（归属 DL_Process，防护门审计状态）
 *----------------------------------------------------------------------------*)
TYPE E_DL_GuardAuditState :
(
    eNormal    := 0,    // 正常：门关、批次可运行 / Normal, door closed
    eHolding   := 10,   // 保持中：批次锁定并记审计 / Holding, batch locked and audited
    eHeld      := 20,   // 已保持：等门关 + 人工确认 / Held, waiting for close plus confirmation
    eResuming  := 30,   // 恢复核实中 / Resuming, residual verification
    eViolation := 40    // 违规：开门超时锁存，需权限复位 / Violation latched, privileged reset required
);
END_TYPE

(*-----------------------------------------------------------------------------
 * 枚举: E_DL_GuardErr（归属 DL_Process，与 FB_DL_MachineGuardAudit 同文件）
 *----------------------------------------------------------------------------*)
TYPE E_DL_GuardErr :
(
    eStNormal   := 16#0005_042B,   // NORMAL / Normal
    eStHolding  := 16#0005_042C,   // HOLDING（批次已锁）/ Holding, batch locked
    eStHeld     := 16#0005_042D,   // HELD（等待恢复确认）/ Held, waiting for confirmation
    eStViolation:= 16#0005_042E,   // VIOLATION（超时锁存）/ Violation latched
    eStResuming := 16#0005_042F    // RESUMING（恢复核实）/ Resuming
);
END_TYPE

(*==============================================================================
 * 功能块: FB_DL_MachineGuardAudit
 * 调用约定: 每个扫描周期无条件调用一次；审计时间戳由上层按任务时基另行记录。
 *============================================================================*)
FUNCTION_BLOCK FB_DL_MachineGuardAudit
VAR_INPUT
    bGuardOpen    : BOOL;                 // 门开信号（TRUE = 门开）/ Guard open signal, TRUE means open
    bBatchActive  : BOOL;                 // 批次运行中 / Batch running
    sOperId       : STRING(32);           // 操作员标识（审计与复位权限）/ Operator identifier for audit and reset
    tMaxOpen      : TIME := T#300S;       // 最长开门时长 [秒]，默认 300 / Maximum open time [s]
    bManualConfirm: BOOL;                 // 人工确认（恢复核实用）/ Manual confirmation for resuming
    bReset        : BOOL;                 // 违规复位请求（上升沿，需操作员标识）/ Violation reset request, edge
END_VAR
VAR_OUTPUT
    eState        : E_DL_GuardAuditState; // 审计状态机当前状态 / Audit state
    bLockBatch    : BOOL;                 // 批次锁定输出 / Batch lock output
    uOpenCnt      : UDINT;                // 开门次数（审计计数，饱和）/ Door-open count, saturating
    sLastOper     : STRING(32);           // 最近一次审计关联操作员 / Last audited operator
    eErr          : E_DL_GuardErr;        // 错误码 / Error code
END_VAR
VAR
    fbGuardTrig   : R_TRIG;               // 门开上升沿实例（无条件调用）/ Guard-open edge instance
    fbResetTrig   : R_TRIG;               // 复位上升沿实例（无条件调用）/ Reset edge instance
    tonOpen       : TON;                  // 开门时长计时器（无条件调用）/ Door-open duration timer
    bOpenPrev     : BOOL;                 // 上拍门信号快照（保守处置参考）/ Previous door signal snapshot
END_VAR
VAR CONSTANT
    DL_GAD_CNT_SAT : UDINT := 16#FFFF_FFFE;   // 开门计数饱和值 [次] / Open count saturation [pcs]
END_VAR

(*------------------------------------------------------------------------------
 * 段 1｜沿检测/TON 每周期无条件调用（仅输入条件化）：超时用状态判定
 *----------------------------------------------------------------------------*)
fbGuardTrig(CLK := bGuardOpen);                        // 门开沿检测无条件刷新 / guard edge refreshed unconditionally
fbResetTrig(CLK := bReset);                            // 复位沿检测无条件刷新 / reset edge refreshed unconditionally
tonOpen(IN := bGuardOpen AND ((eState = E_DL_GuardAuditState.eHolding)
                           OR (eState = E_DL_GuardAuditState.eHeld)), PT := tMaxOpen);   // 开门时长计时 / open-duration timing
bOpenPrev := bGuardOpen;                               // 门信号快照推进 / snapshot advanced

(*------------------------------------------------------------------------------
 * 段 2｜违规复位：需操作员标识非空（权限侧要求，空标识一律拒绝）
 *----------------------------------------------------------------------------*)
IF fbResetTrig.Q AND (eState = E_DL_GuardAuditState.eViolation) THEN
    IF sOperId <> '' THEN                              // 标识非空才允许复位 / non-empty operator required
        eState := E_DL_GuardAuditState.eNormal;        // 解锁回正常 / back to normal
        bLockBatch := FALSE;                           // 批次解锁 / batch unlocked
    END_IF
    // 空标识：保持 VIOLATION 锁存（权限复位不在本块裁决）/ empty id keeps the violation latched
END_IF

(*------------------------------------------------------------------------------
 * 段 3｜门开上升沿：批次活动中 → HOLDING（锁批次 + 审计）；否则保守置 Held
 *----------------------------------------------------------------------------*)
IF fbGuardTrig.Q THEN
    IF uOpenCnt < DL_GAD_CNT_SAT THEN
        uOpenCnt := uOpenCnt + 1;                      // 开门次数饱和自增 [次] / saturating open count
    END_IF
    sLastOper := sOperId;                              // 审计操作员留痕 / operator audited
    IF bBatchActive THEN
        eState := E_DL_GuardAuditState.eHolding;       // 批次活动：HOLDING / batch active: holding
        bLockBatch := TRUE;                            // 锁批次 / batch locked
    ELSE
        eState := E_DL_GuardAuditState.eHeld;          // 无批次：直接 Held（无需锁）/ no batch: held directly
        bLockBatch := TRUE;                            // 保守侧仍锁批次（防误运行）/ conservatively locked
    END_IF
END_IF

(*------------------------------------------------------------------------------
 * 段 4｜审计状态机：CASE 含 ELSE 兜底（ELSE → VIOLATION 锁存）
 *----------------------------------------------------------------------------*)
CASE eState OF

    E_DL_GuardAuditState.eNormal:
        bLockBatch := FALSE;                           // 正常：批次不锁 / batch unlocked
        eErr := E_DL_GuardErr.eStNormal;               // 码 042B / code normal

    E_DL_GuardAuditState.eHolding:
        bLockBatch := TRUE;                            // 保持中：批次锁 / batch locked
        eErr := E_DL_GuardErr.eStHolding;              // 码 042C / code holding
        eState := E_DL_GuardAuditState.eHeld;          // 审计记录完成：进 Held / audit recorded, enter held

    E_DL_GuardAuditState.eHeld:
        bLockBatch := TRUE;                            // 已保持：批次锁 / batch locked
        eErr := E_DL_GuardErr.eStHeld;                 // 码 042D / code held
        IF (NOT bGuardOpen) AND bManualConfirm THEN
            eState := E_DL_GuardAuditState.eResuming;  // 门关 + 人工确认：进核实 / closed plus confirmed: resuming
        ELSIF tonOpen.Q THEN
            eState := E_DL_GuardAuditState.eViolation; // 开门超时：违规锁存 / open timeout: violation latch
            bLockBatch := TRUE;                        // 违规：批次锁保持 / lock held
        END_IF

    E_DL_GuardAuditState.eResuming:
        bLockBatch := TRUE;                            // 核实中：批次锁保持（未核实不放行）/ lock held while verifying
        eErr := E_DL_GuardErr.eStResuming;             // 码 042F / code resuming
        IF (NOT bGuardOpen) AND bManualConfirm THEN
            eState := E_DL_GuardAuditState.eNormal;    // 核实通过（无残留）：回正常 / verified: back to normal
            bLockBatch := FALSE;                       // 批次解锁 / batch unlocked
        ELSIF tonOpen.Q THEN
            eState := E_DL_GuardAuditState.eViolation; // 核实期开门超时：违规锁存 / timeout while verifying: violation
        END_IF

    E_DL_GuardAuditState.eViolation:
        bLockBatch := TRUE;                            // 违规：批次锁保持（需权限复位）/ lock held, privileged reset only
        eErr := E_DL_GuardErr.eStViolation;            // 码 042E / code violation

    ELSE
        eState := E_DL_GuardAuditState.eViolation;     // 非法状态兜底：按违规锁存（保守侧）/ illegal-state fallback to violation
        bLockBatch := TRUE;                            // 批次锁保持 / lock held
        eErr := E_DL_GuardErr.eStViolation;            // 兜底码（违规段，反证句：输出同为锁批次+锁存）/ fallback code

END_CASE
END_FUNCTION_BLOCK

(* ---- FB_DL_MakeupWaterDosing.st ---- *)
(*
  Name        : FB_DL_MakeupWaterDosing
  Category    : DL_Process
  Version     : 1.0.0
  Purpose     : 补水定量加药：累计补水流量体积，每到设定批量体积即触发一次定比投加（加药量 = 批量 × 投加比），投加脉冲单拍输出并累计批次数；/ Makeup-water proportional dosing: accumulate makeup volume and trigger one proportional dose (dose = batch x ratio) each time the batch volume is reached, with a single-scan dose pulse and batch count
  溯源        : ROADMAP L501（未勾真缺口），IEC 61131-3 标准语义的道莅防御性实现
  Boundary    : ① 组态闸：批量体积/投加比/采样周期任一非正 → 锁存故障；
                ② 体积换算：m³/h → L/s 除子 3.6 为常量，无组态除零风险；采样周期正域由组态闸保证；
                ③ 单次只结算一个批次（净额单点写入），剩余体积保留进位（大流量不丢批）；
                ④ 投加脉冲为单拍（内部置位 → 出口统一映射，R187），批次数饱和累加；
                ⑤ 负流量（回流）不计入累计，防倒吸误触发。
*)
TYPE E_DL_MwdState :
(
    eIdle  := 0,                             (* 未使能 / Disabled *)
    eAcc   := 10,                            (* 体积累计 / Accumulating *)
    eFault := 90                             (* 故障锁存相 / Fault latched *)
);
END_TYPE

TYPE E_DL_MwdCause :
(
    eNone       := 0,                        (* 无故障成因 / No cause *)
    eCfgIllegal := 1,                        (* 组态非法：批量/比值/周期越域 / Illegal config *)
    ePhaseBad   := 2                         (* 非法相位兜底 / Illegal phase fallback *)
);
END_TYPE

FUNCTION_BLOCK FB_DL_MakeupWaterDosing
VAR_INPUT
    fFlowNow  : REAL := 0.0;                 (* 补水瞬时流量（负值为回流），[m³/h] / Makeup flow, negative = backflow *)
    fBatchVol : REAL := 100.0;               (* 触发批量体积，域 > 0 [L] / Batch volume trigger, > 0 *)
    fDoseRatio: REAL := 0.5;                 (* 投加比（加药量/补水体积），域 > 0 [L/m³] / Dose ratio, > 0 *)
    tSample   : TIME := T#100MS;             (* 采样周期，域 > T#0S [ms] / Sampling period, > 0 *)
    bEnable   : BOOL := TRUE;                (* 使能 [-] / Enable *)
    bReset    : BOOL := FALSE;               (* 复位命令，上升沿清累计与批次 [-] / Reset command *)
END_VAR
VAR_OUTPUT
    fVolAcc   : REAL;                        (* 当前批次已累计体积 [L] / Volume accumulated in current batch *)
    fVolTotal : REAL;                        (* 累计补水总量（生命周期）[L] / Lifetime accumulated volume *)
    fDoseVol  : REAL;                        (* 本次投加量（脉冲拍有效）[L] / Dose volume of this pulse *)
    bDosePulse: BOOL;                        (* 投加触发单拍脉冲 [-] / Dose trigger single-scan pulse *)
    nBatchCnt : UDINT;                       (* 已完成批次数（饱和）[批] / Completed batches, saturated *)
    eState    : E_DL_MwdState;               (* 状态出口 / State outlet *)
    eCause    : E_DL_MwdCause;               (* 故障成因出口（R190 归因唯一） / Fault cause outlet *)
    bError    : BOOL;                        (* 故障锁存标志 [-] / Fault latch flag *)
END_VAR
VAR
    _eState  : E_DL_MwdState := E_DL_MwdState.eIdle;     (* 内部相位（CASE 唯一写入目标） / Internal phase *)
    _eCause  : E_DL_MwdCause := E_DL_MwdCause.eNone;     (* 故障成因锁存量 / Latched cause *)
    rtReset  : R_TRIG;                       (* 复位沿实例，段 0 无条件调用 / Reset edge instance *)
    _bFault  : BOOL;                         (* 故障锁存位 / Latched fault bit *)
    _bCfgBad : BOOL;                         (* 组态非法当拍量 / Illegal config this scan *)
    _bFinite : BOOL;                         (* 输入有限性当拍量 / Input finiteness *)
    _bDoseC  : BOOL;                         (* 投加脉冲内部单拍量（出口统一映射） / Dose internal pulse *)
    _fDtSec  : REAL;                         (* 采样周期秒值 [s] / Period in seconds *)
    _fDvL     : REAL;                        (* 本拍补水体积增量 [L] / Volume increment this scan *)
    _fAcc    : REAL;                         (* 批次累计内部量 [L] / Batch accumulator *)
    _fTotal  : REAL;                         (* 生命周期累计内部量 [L] / Lifetime accumulator *)
    _fDose   : REAL;                         (* 本次投加量计算值 [L] / Dose calculation *)
    _fZero   : REAL;                         (* 实数零常量 [-] / Zero constant *)
END_VAR
VAR CONSTANT
    DL_MWD_EPS    : REAL  := 1.0E-6;         (* 判零容差 [-] / Epsilon *)
    DL_MWD_M3H2LS : REAL  := 3.6;            (* m³/h → L/s 换算常量（1 m³/h = 1/3.6 L/s）[-] / Conversion constant *)
    DL_MWD_CNTMAX : UDINT := 4294967295;     (* 批次数饱和上限（R28）[批] / Batch count cap *)
END_VAR

(* —— 段 0：当拍判据派生 + 实例无条件刷新（R228A） —— *)
_fDtSec := TIME_TO_LREAL(tSample) / 1000.0;                                    (* 周期秒化（除子常量 1000） / Period to seconds *)
_bCfgBad := (fBatchVol <= DL_MWD_EPS)                                          (* 批量体积正域闸 / Batch volume gate *)
            OR (fDoseRatio <= DL_MWD_EPS)                                      (* 投加比正域闸 / Dose ratio gate *)
            OR NOT (tSample > T#0S);                                           (* 采样周期正域闸 / Period gate *)
rtReset(CLK := bReset);                                                        (* 复位沿每拍必调 / Reset edge every scan *)
_bFinite := (fFlowNow = fFlowNow) AND ((fFlowNow - fFlowNow) = (fFlowNow - fFlowNow));   (* NaN 自反 + Inf 差判 / NaN and Inf gate *)
_fZero := 0.0;                                                                 (* 零常量装载 / Zero constant load *)

(* —— 段 1：单拍量预清零（R107） —— *)
_bDoseC := FALSE;                                                              (* 投加脉冲内部量预清 / Dose preset *)
fDoseVol := 0.0;                                                               (* 投加量出口预清（脉冲拍外恒 0） / Dose outlet preset *)

(* —— 段 2：复位沿处理（作用域：清故障 + 清累计 + 清批次 + 迁 eIdle，R283 逐项声明） —— *)
IF rtReset.Q THEN
    _bFault := FALSE;                                                          (* 清故障锁存 / Clear fault *)
    _eCause := E_DL_MwdCause.eNone;                                            (* 清成因 / Clear cause *)
    _fAcc := 0.0;                                                              (* 清批次累计 / Clear batch accumulator *)
    _fTotal := 0.0;                                                            (* 清总量累计 / Clear lifetime accumulator *)
    fVolAcc := 0.0;                                                            (* 清批次出口 / Clear batch outlet *)
    fVolTotal := 0.0;                                                          (* 清总量出口 / Clear total outlet *)
    nBatchCnt := 0;                                                            (* 清批次数 / Clear batch count *)
    _eState := E_DL_MwdState.eIdle;                                            (* 迁未使能相 / Back to idle *)
END_IF

(* —— 段 3：组态故障锁存（锁存至复位沿，R189） —— *)
IF _bCfgBad AND NOT _bFault THEN
    _bFault := TRUE;                                                           (* 锁存故障位 / Latch fault *)
    _eCause := E_DL_MwdCause.eCfgIllegal;                                      (* 成因：组态非法 / Cause: illegal config *)
    _eState := E_DL_MwdState.eFault;                                           (* 同步迁故障相 / Migrate to fault *)
END_IF

(* —— 段 4：CASE 主状态机（ELSE 兜底迁 eFault，红线 6） —— *)
CASE _eState OF
    E_DL_MwdState.eIdle:                                                       (* 未使能：不累计 / Disabled *)
        fVolAcc := _fAcc;                                                      (* 出口镜像（保持当前批次进度） / Outlet mirror *)
        fVolTotal := _fTotal;                                                  (* 总量出口镜像 / Total outlet mirror *)
        IF bEnable AND NOT _bFault THEN
            _eState := E_DL_MwdState.eAcc;                                     (* 使能进入累计 / Enter accumulating *)
        END_IF
    E_DL_MwdState.eAcc:                                                        (* 累计相：体积积分 + 批量触发 / Accumulating *)
        IF NOT bEnable THEN
            _eState := E_DL_MwdState.eIdle;                                    (* 失能回未使能 / Back to idle *)
        ELSIF _bFinite AND (_fDtSec > DL_MWD_EPS) THEN
            _fDvL := fFlowNow / DL_MWD_M3H2LS * _fDtSec;                       (* 体积增量 = (m³/h→L/s)·s（除子常量）[L] / Volume increment *)
            IF _fDvL > _fZero THEN                                             (* 负流量（回流）不计入（边界⑤） / Backflow ignored *)
                _fAcc := _fAcc + _fDvL;                                        (* 批次累计 / Batch accumulate *)
                _fTotal := _fTotal + _fDvL;                                    (* 总量累计 / Lifetime accumulate *)
            END_IF
            IF _fAcc >= fBatchVol THEN                                         (* 到批量：触发一次投加 / Batch reached: dose once *)
                _fDose := fBatchVol * fDoseRatio;                              (* 投加量 = 批量 × 比值 [L] / Dose volume *)
                fDoseVol := _fDose;                                            (* 投加量出口（脉冲拍有效） / Dose outlet *)
                _bDoseC := TRUE;                                               (* 脉冲内部置位（出口统一映射，R187） / Pulse internal *)
                _fAcc := _fAcc - fBatchVol;                                    (* 剩余体积进位，不丢批（净额单点写入） / Carry remainder *)
                IF _fAcc < _fZero THEN
                    _fAcc := _fZero;                                           (* 进位后下限保护（浮点舍入） / Carry floor *)
                END_IF
                IF nBatchCnt < DL_MWD_CNTMAX THEN
                    nBatchCnt := nBatchCnt + 1;                                (* 批次净额 +1（同拍不叠加） / Net +1 *)
                END_IF
            END_IF
            fVolAcc := _fAcc;                                                  (* 批次进度出口 / Batch progress outlet *)
            fVolTotal := _fTotal;                                              (* 总量出口 / Total outlet *)
        END_IF                                                                 (* 非有限输入：本拍不累计 / Non-finite: skip *)
    E_DL_MwdState.eFault:                                                      (* 故障相：冻结保持末值，仅复位沿出 / Fault *)
        ;                                                                      (* 锁存回放（R28） / Replay from latch *)
    ELSE                                                                       (* 非法相位兜底迁安全态 / Illegal phase fallback *)
        _eState := E_DL_MwdState.eFault;                                       (* 迁故障相 / To fault *)
        _bFault := TRUE;                                                       (* 同步锁存 / Latch *)
        _eCause := E_DL_MwdCause.ePhaseBad;                                    (* 成因：非法相位 / Cause: illegal phase *)
END_CASE

(* —— 段 5：出口映射（内部 _b* → 输出单拍，R187；名实双出口，R191） —— *)
bDosePulse := _bDoseC;                                                         (* 投加脉冲单拍出口 / Dose pulse outlet *)
bError := _bFault;                                                             (* 故障标志镜像 / Fault flag mirror *)
eState := _eState;                                                             (* 状态出口 / State outlet *)
eCause := _eCause;                                                             (* 成因出口 / Cause outlet *)
END_FUNCTION_BLOCK

(* ---- FB_DL_MaterialHoldTimeEnforce.st ---- *)
(*
  ==================================================================
  组件名 Component  : FB_DL_MaterialHoldTimeEnforce
  分类   Category   : DL_Process
  复杂度 Complexity  : cx5
  版本   Version    : 1.0.0
  功能   Purpose    : 物料保持时限强制。批次开始沿起累计保持时长，超时限判
                      NG 锁存（ISA-88 批次语境）；复检合格沿解锁放行并出
                      单拍放行脉冲；批次与超时台账计数出口。GMP 保持时限
                      公开语义（中间品 / 批次在制时限管理）。
  来源   Source     : self（GMP 保持时限公开语义，ISA-88 批次语境次源）
  溯源   Origin     : IEC 61131-3 标准语义的道莅防御性实现；保持时限与复检
                      放行为行业公开流程语义，clean-room 自研实现，未复制
                      任何厂商私有库源码。
  平台   Platform   : 纯 IEC 61131-3（Standard.library: R_TRIG / F_TRIG，无私有库）
  分工声明 Split     : 与 DL_Process 存量批次追溯件（批次履历类）分工——履历
                      件做批次数据记录，本件只做保持时限判定与放行门控；
                      不做配方切换与批次数据缓存。
  作者   Author     : 道莅代码库 · PLC 编程专家（R58）
  ------------------------------------------------------------------
  边界 Boundary     :
                      一 代理量三句声明（R95）：fScanPeriodMin 为每次调用的
                         代表时长（代理值）；覆盖任务周期 0.1..10 分钟调用
                         节拍；覆盖不到的区间（调用节拍外事件）由调用方批
                         次信号沿精度兜尾；
                      二 组态域：fHoldLimitMin > 0 且非有限、fScanPeriodMin
                         > 0 且非有限；越域锁存（解除 = bReset 沿，R188）；
                      三 超时 NG 锁存解除路径 = bRecheckOk 上升沿（复检放行，
                         唯一路径，R188 头注释声明）；放行脉冲为单拍（R25：
                         预清零点在段 3，置位点在段 5，两段式映射）；
                      四 复位沿作用域：清故障锁存 / 清台账计数 / 清保持累计
                         与锁存（三项逐项声明）；
                      五 无全局变量、无外部变量声明、无物理地址寻址。
  修订记录 Revision  :
    2026-11-21  v1.0.0  R58 首版（批 4 · 序号 15）
  ==================================================================
*)

FUNCTION_BLOCK FB_DL_MaterialHoldTimeEnforce
VAR_INPUT
    bEnable        : BOOL := TRUE;   // 使能，失能冻结判定（输出保持）[-] / enable, disabling freezes the verdicts
    bReset         : BOOL := FALSE;  // 复位上升沿清锁存与台账 [-] / reset rising edge clears the latch and the ledger
    bBatchStart    : BOOL := FALSE;  // 批次开始信号（沿生效）[-] / the batch start signal, edge effective
    bBatchActive   : BOOL := FALSE;  // 批次在制电平 [-] / the batch active level
    bRecheckOk     : BOOL := FALSE;  // 复检合格信号（沿生效）[-] / the recheck pass signal, edge effective
    fHoldLimitMin  : LREAL := 120.0; // 保持时限 [分钟]，域 大于 0 / the hold limit [minute], above zero
    fScanPeriodMin : LREAL := 1.0;   // 每次调用的代表时长 [分钟]（代理量，边界一）/ the representative duration per call [minute]
END_VAR
VAR_OUTPUT
    bExpired        : BOOL := FALSE; // 超时限 NG 锁存出口 [-] / the expired NG latch outlet
    bReleaseOk      : BOOL := FALSE; // 复检放行单拍出口 [-] / the recheck release pulse outlet
    fHoldElapsedMin : LREAL := 0.0;  // 已保持时长出口 [分钟] / the elapsed hold duration outlet [minute]
    nBatchCnt       : UDINT := 0;    // 累计批次数 [批] / the total batch count [batch]
    nExpiredCnt     : UDINT := 0;    // 超时批次数 [批] / the expired batch count [batch]
    bError          : BOOL := FALSE; // 域闸故障锁存标志 [-] / the domain gate fault latch flag
END_VAR
VAR
    rtStart : R_TRIG; // 批次开始沿检测，段 0 无条件刷新 / the batch start edge
    rtRel   : R_TRIG; // 复检合格沿检测，段 0 无条件刷新 / the recheck edge
    ftBatch : F_TRIG; // 批次结束沿检测（在制下降沿），段 0 无条件刷新 / the batch end edge, a falling edge
    rtReset : R_TRIG; // 复位沿检测，段 0 无条件刷新 / the reset edge
    _bCnt   : BOOL := FALSE; // 保持计时进行中 [-] / the hold timing active
    _bExpL  : BOOL := FALSE; // 超时 NG 锁存位（解除 = 复检合格沿）/ the expired NG latch bit
    _bRel   : BOOL := FALSE; // 放行脉冲内部保持量（统一出口映射单拍）/ the release pulse internal holder
    _bLatch : BOOL := FALSE; // 域闸故障锁存位 [-] / the domain gate latch bit
    _bInit  : BOOL := FALSE; // 首扫初始化完成标志（R310）/ the first scan flag
END_VAR
VAR CONSTANT
    DL_MHT_CNTMAX : UDINT := 4294967294; // 台账计数钳定界 [批]，防 UDINT 回绕 / the ledger clamp against a wrap
END_VAR

// 段 0｜沿检测无条件周期刷新（禁入分支，FB50-1）/ segment 0, the unconditional refresh
rtStart(CLK := bBatchStart); // 批次开始沿 / the batch start edge
rtRel(CLK := bRecheckOk); // 复检合格沿 / the recheck edge
ftBatch(CLK := bBatchActive); // 批次结束沿 / the batch end edge
rtReset(CLK := bReset); // 复位沿 / the reset edge

// 段 1｜首扫初始化（R310）/ segment 1, the first scan
IF NOT _bInit THEN // 首扫一拍 / the first scan
    _bInit := TRUE; // 置首扫标志 / raise the flag
END_IF

// 段 2｜复位沿作用域：清故障锁存 / 清台账 / 清保持累计与锁存（三项逐项声明，边界四）/ segment 2, the reset edge scope
IF rtReset.Q THEN // 复位沿 / the reset edge
    _bLatch := FALSE; // 作用域一：清域闸锁存 / scope one, clear the latch
    _bExpL := FALSE; // 作用域一：清 NG 锁存（复位沿为 NG 锁存的辅助解除路径）/ scope one, clear the NG latch
    nBatchCnt := 0; // 作用域二：清批次台账 / scope two, clear the batch ledger
    nExpiredCnt := 0; // 作用域二：清超时台账 / scope two, clear the expired ledger
    fHoldElapsedMin := 0.0; // 作用域三：清保持累计 / scope three, clear the hold accumulator
    _bCnt := FALSE; // 作用域三：清计时进行 / scope three, clear the timing
END_IF

// 段 3｜组态域闸 + 单拍标志预清零（R25）/ segment 3, the config gate and the single shot presets
IF (fHoldLimitMin <> fHoldLimitMin) OR ((fHoldLimitMin - fHoldLimitMin) <> (fHoldLimitMin - fHoldLimitMin)) // 时限非有限 / a non finite limit
OR (fHoldLimitMin <= 0.0) // 时限域 / the limit domain
OR (fScanPeriodMin <> fScanPeriodMin) OR ((fScanPeriodMin - fScanPeriodMin) <> (fScanPeriodMin - fScanPeriodMin)) // 代理周期非有限 / a non finite period
OR (fScanPeriodMin <= 0.0) THEN // 代理周期域 / the period domain
    IF NOT _bLatch THEN // 未锁存才置位 / latch only while unlatched
        _bLatch := TRUE; // 置域闸锁存 / raise the latch
    END_IF
END_IF
bError := _bLatch; // 故障标志与锁存位同源（R191 名实双出口）/ the flag shares the latch
bReleaseOk := FALSE; // 放行单拍每拍预清零（R25，置位点在段 5 统一出口）/ the release pulse preset false each scan

// 段 4｜批次受理与保持累计（域内才推进，边界一二）/ segment 4, the batch admission and the hold accumulation
IF (rtStart.Q OR (bBatchActive AND (NOT _bCnt) AND (NOT _bExpL))) AND (NOT _bLatch) THEN // 批次开始沿或在制重新受理 / a batch start edge or a re admission
    IF rtStart.Q THEN // 仅开始沿计台账 / only the start edge counts the ledger
        IF nBatchCnt < DL_MHT_CNTMAX THEN // 台账防回绕 / the ledger wrap guard
            nBatchCnt := nBatchCnt + 1; // 批次计数推进 / advance the batch count
        END_IF
    END_IF
    fHoldElapsedMin := 0.0; // 保持累计清零起算 / clear the accumulator
    _bCnt := TRUE; // 启动保持计时 / start the timing
    _bExpL := FALSE; // 新批次清 NG 锁存（换批自动解锁声明）/ clear the NG latch on a new batch
END_IF
IF _bCnt AND bBatchActive AND (NOT _bLatch) THEN // 计时中且在制且域内 / while timing, active, inside the domain
    fHoldElapsedMin := fHoldElapsedMin + fScanPeriodMin; // 保持累计推进（代理量，边界一）/ advance the accumulator
    IF (fHoldElapsedMin > fHoldLimitMin) AND (NOT _bExpL) THEN // 首次越限（单批只计一次台账）/ the first overrun, one ledger entry per batch
        _bExpL := TRUE; // 置 NG 锁存 / raise the NG latch
        IF nExpiredCnt < DL_MHT_CNTMAX THEN // 台账防回绕 / the ledger wrap guard
            nExpiredCnt := nExpiredCnt + 1; // 超时计数推进 / advance the expired count
        END_IF
    END_IF
END_IF
IF ftBatch.Q THEN // 批次结束沿（在制下降）/ a batch end edge
    _bCnt := FALSE; // 停止计时（累计量保留供显示）/ stop the timing, the accumulator retained
END_IF

// 段 5｜复检放行与统一出口（边界三）/ segment 5, the release and the unified outlet
IF _bExpL AND rtRel.Q THEN // NG 锁存且复检合格沿（解除路径，R188）/ the NG latch with the recheck edge
    _bExpL := FALSE; // 解除 NG 锁存 / release the NG latch
    _bRel := TRUE; // 置放行内部保持量 / raise the release holder
END_IF
bExpired := _bExpL; // NG 锁存出口单点映射 / the NG outlet mapped
IF _bRel THEN // 放行内部保持量 → 统一出口单拍映射（两段式，R189）/ the holder mapped to the pulse
    bReleaseOk := TRUE; // 放行单拍 / the release pulse
    _bRel := FALSE; // 消费保持量 / consume the holder
END_IF
END_FUNCTION_BLOCK

(* ---- FB_DL_MercerCausticConcWatch.st ---- *)
(*
  Name: FB_DL_MercerCausticConcWatch
  Category: DL_Process
  Version: 1.0.0
  Round: R91 / 2026-11-25
  开源溯源：clean-room 自研（族 间歇式溢流染色与丝光整理，ST 开源生态实测 0 命中，无外部代码引入）
  功能：1) 丝光碱浓度双向监视，超限判据各自去抖后锁存：
           低于 fConcLoGpl 进低浓相并置补碱请求（xMakeupReq），丝光不足会导致纤维膨化不够；
           高于 fConcHiGpl 进高浓相并置稀释请求（xDiluteReq），碱浓过高会损伤纤维并增加中和负荷。
        2) 连续失效计数：每次「去抖确认的越限」使 nFailCount 加一，回到带内即清零；
           计数达到 fFailMax（INT 引脚）时升级为故障锁存（码 0415）——
           这是「反复越限、补液联动无效」的累积证据，比单次越限更值得停机处理。
        3) 三级语义：带内正常（信息级码 0414）→ 越限锁存（故障级 0412 / 0413）→ 累计失效（0415）。
           任一故障级锁存均不直接停设备，由上层决定是否停止进布（本件只监视不驱动工艺阀）。
  边界条件：1) 非有限值闸：浓度与两个阈值先过 NOT(x > -DL_BIG AND x < DL_BIG)，同时拦 NaN 与 Inf；
           命中即锁码 0417 进故障相 —— 绝不把 NaN 拿去与浓度阈比较
           （NaN 比较恒假会把「碱浓电极断线」伪装成「浓度正常」，R19）。
        2) 阈值域闸：须满足 0.0 < fConcLoGpl < fConcHiGpl <= DL_CONC_HI，越域锁码 0417
           （两级判据重叠会让某向永不触发）；tDebounce 必须 > T#0S（零窗使判据无滞后直达停机）。
        3) 计数域闸：fFailMax 必须 >= 1（为 0 会使累计判据恒真，一上电就报 0415）。
        4) 浓度量级闸：实测浓度须落在 [0.0, DL_CONC_HI] 内，越域锁码 0417（电极标定丢失）。
        5) 定时器周期刷新（R7）：两个去抖 TON 与复位边沿全部在 CASE 之外无条件调用。
        6) 故障解除路径：低浓/高浓相内 xReset 上升沿即清锁存回正常（可达）；
           故障相内还必须同时满足 NOT xFault 且入参/组态合法才可解除（不自恢复）。
        7) 状态机兜底：CASE 全态覆盖 + ELSE 强制回故障相并置码 0418、清全部输出。
        8) 输出安全初值（R25）：两个报警位、两个请求位初值 FALSE，nFailCount 初值 0，
           正常相显式赋值，防「上电未初始化直穿」。
  量纲自证：fConcGpl 与 fConcLoGpl / fConcHiGpl 全为质量浓度 [g/L]，比较两侧同量纲；
           nFailCount / fFailMax 为计数 [count]，无因次。
  码表 Error codes（本件子带 0091_041x，故障级一律 3 行内置 _uFault/_bFault/_eState）:
    16#0091_0411 信息级：碱浓度接近下限，尚在去抖窗内（不置故障位）
    16#0091_0412 故障级：碱浓度低于下限（去抖确认，请求补碱）
    16#0091_0413 故障级：碱浓度高于上限（去抖确认，请求稀释）
    16#0091_0414 信息级：碱浓度在工艺带内（不置故障位）
    16#0091_0415 故障级：连续失效计数达上限（补液联动无效）
    16#0091_0416 故障级：外部故障输入 xFault
    16#0091_0417 故障级：入参非有限，或阈值/计数/去抖窗组态越域
    16#0091_0418 故障级：状态机落 ELSE 兜底（非法相位 ID）

  修订历史 Revision :
    2026-11-25  v1.0.0  R91 首版
*)

TYPE E_DL_JbsCausticConcState :
(
    eJbsConcNormal := 0,    // 正常：浓度在工艺带内 / Normal, concentration within the process band
    eJbsConcLow    := 10,   // 低浓：去抖确认后锁存，请求补碱 / Low, latched after debounce, make-up requested
    eJbsConcHigh   := 20,   // 高浓：去抖确认后锁存，请求稀释 / High, latched after debounce, dilution requested
    eJbsConcFault  := 90    // 故障：入参/组态非法或累计失效，锁存待解除 / Fault, invalid input or repeated failures
);
END_TYPE

FUNCTION_BLOCK FB_DL_MercerCausticConcWatch
VAR_INPUT
    xEnable      : BOOL;    // 监视使能 [bool] / Monitoring enable [bool]
    xReset       : BOOL;    // 报警/故障复位（上升沿有效）[bool] / Alarm and fault reset, rising edge [bool]
    xFault       : BOOL;    // 外部故障汇总 [bool] / External fault aggregate [bool]
    fConcGpl     : REAL;    // 实测碱质量浓度 [g/L] / Measured caustic concentration [g/L]
    fConcLoGpl   : REAL;    // 浓度工艺下限 [g/L] / Concentration process low limit [g/L]
    fConcHiGpl   : REAL;    // 浓度工艺上限 [g/L] / Concentration process high limit [g/L]
    tDebounce    : TIME;    // 判据去抖窗 [TIME] / Criteria debounce window [TIME]
    fFailMax     : INT;     // 连续失效计数上限 [count] / Consecutive failure count limit [count]
END_VAR
VAR_OUTPUT
    xLowAlarm    : BOOL;    // 低浓报警（锁存）[bool] / Low concentration alarm, latched [bool]
    xHighAlarm   : BOOL;    // 高浓报警（锁存）[bool] / High concentration alarm, latched [bool]
    xMakeupReq   : BOOL;    // 补碱（补液）联动请求 [bool] / Caustic make-up request [bool]
    xDiluteReq   : BOOL;    // 稀释（补水）联动请求 [bool] / Dilution water request [bool]
    nFailCount   : INT;     // 连续失效计数 [count] / Consecutive failure count [count]
    eState       : E_DL_JbsCausticConcState;   // 状态出口，段尾单点映射 / State outlet, single-point mapped
    nErrId       : UDINT;   // 事件码，0 = 无事件 / Event code, 0 = none
END_VAR
VAR
    tonLow       : TON;     // 低浓去抖定时 [TIME] / Low concentration debounce timer
    tonHigh      : TON;     // 高浓去抖定时 [TIME] / High concentration debounce timer
    rtReset      : R_TRIG;  // 复位上升沿检测 [bool] / Reset rising edge detector
    _eState      : E_DL_JbsCausticConcState := E_DL_JbsCausticConcState.eJbsConcNormal;   // 内部相位（CASE 唯一写入目标）
    _iFailCnt    : INT := 0;        // 内部连续失效计数 [count] / Internal consecutive failure count [count]
    _bFinOk      : BOOL := FALSE;   // 实值入参有限性总闸结果 / Finiteness gate aggregate result
    _bCfgOk      : BOOL := FALSE;   // 阈值与计数组态域闸结果 / Threshold and count domain gate result
    _bLowRaw     : BOOL := FALSE;   // 低浓原始判据 [bool] / Raw low concentration criterion
    _bHighRaw    : BOOL := FALSE;   // 高浓原始判据 [bool] / Raw high concentration criterion
    _bLowL       : BOOL := FALSE;   // 低浓锁存位 [bool] / Latched low alarm flag
    _bHighL      : BOOL := FALSE;   // 高浓锁存位 [bool] / Latched high alarm flag
    _bFault      : BOOL := FALSE;   // 故障锁存位 [bool] / Latched fault flag
    _uInfo       : UDINT := 16#0000_0000;   // 信息码，每拍重算 / Info code, recomputed every cycle
    _uFault      : UDINT := 16#0000_0000;   // 故障码锁存 / Latched fault code
END_VAR
VAR CONSTANT
    DL_EPS       : REAL := 1.0E-9;      // 数值零闸阈值 [-] / Numeric zero gate threshold [-]
    DL_BIG       : REAL := 1.0E12;      // 非有限值闸量级上限 [-] / Finiteness gate magnitude [-]
    DL_CONC_HI   : REAL := 1000.0;      // 浓度量级闸上限 [g/L] / Concentration magnitude upper bound [g/L]
    DL_CNT_HI    : INT := 10000;        // 计数显示上限 [count] / Count display upper bound [count]
END_VAR

(* —— 段 0：单拍量预清零（锁存量 _uFault/_bFault/_bLowL/_bHighL/_iFailCnt 不入清单，R187①） —— *)
_uInfo := 16#0000_0000;                     // 信息码每拍重算 / Info code recomputed
nErrId := 16#0000_0000;                     // 事件码缺省无事件 / Event code defaults to none

(* —— 段 1：非有限值闸与组态域闸（R19：不拿 NaN 去比较浓度阈） —— *)
_bFinOk := (fConcGpl > -DL_BIG) AND (fConcGpl < DL_BIG)
           AND (fConcLoGpl > -DL_BIG) AND (fConcLoGpl < DL_BIG)
           AND (fConcHiGpl > -DL_BIG) AND (fConcHiGpl < DL_BIG);
_bCfgOk := (fConcLoGpl > DL_EPS)                            // 下限必须为正
           AND (fConcHiGpl > fConcLoGpl)                     // 上限必须严格大于下限
           AND (fConcHiGpl <= DL_CONC_HI)                    // 上限须在量级闸内
           AND (fConcGpl >= 0.0) AND (fConcGpl <= DL_CONC_HI)   // 实测浓度量级闸
           AND (tDebounce > T#0S)                            // 去抖窗必须为正
           AND (fFailMax >= 1);                              // 计数上限至少为 1

(* —— 段 2：原始判据（取未钳制的实测浓度，禁先夹后判，R24） —— *)
_bLowRaw := _bFinOk AND _bCfgOk AND (fConcGpl < fConcLoGpl);             // 低浓原始判据
_bHighRaw := _bFinOk AND _bCfgOk AND (fConcGpl > fConcHiGpl);            // 高浓原始判据

(* —— 段 3：定时器与边沿无条件周期刷新（R7：调用语句不得置于 IF/CASE 内） —— *)
rtReset(CLK := xReset);                                                     // 复位上升沿，每拍必调
tonLow(IN := _bLowRaw AND (NOT _bFault), PT := tDebounce);                  // 低浓去抖
tonHigh(IN := _bHighRaw AND (NOT _bFault), PT := tDebounce);                // 高浓去抖

(* —— 段 4：全局故障拦截（优先级最高；已锁存则不再改写码值，禁同拍抹除） —— *)
IF xFault AND (NOT _bFault) THEN
    _uFault := 16#0091_0416;                // 故障级：外部故障输入
    _bFault := TRUE;                        // 锁存（3 行内置，R45 配对）
    _eState := E_DL_JbsCausticConcState.eJbsConcFault;
END_IF
IF ((NOT _bFinOk) OR (NOT _bCfgOk)) AND (NOT _bFault) THEN
    _uFault := 16#0091_0417;                // 故障级：入参非有限或组态越域（内部成员已分离）
    _bFault := TRUE;                        // 锁存
    _eState := E_DL_JbsCausticConcState.eJbsConcFault;
END_IF

(* —— 段 5：相位机（只做迁移与锁存；出口在段 7 单点映射） —— *)
CASE _eState OF

E_DL_JbsCausticConcState.eJbsConcNormal:
    IF NOT xEnable THEN
        _uInfo := 16#0091_0414;             // 信息级：监视关闭，浓度保持上拍结论（不置故障位）
    ELSIF tonLow.Q THEN
        _uFault := 16#0091_0412;            // 故障级：碱浓度低于下限（去抖确认）
        _bLowL := TRUE;                     // 低浓锁存
        _iFailCnt := _iFailCnt + 1;         // 连续失效计数加一
        _eState := E_DL_JbsCausticConcState.eJbsConcLow;
    ELSIF tonHigh.Q THEN
        _uFault := 16#0091_0413;            // 故障级：碱浓度高于上限（去抖确认）
        _bHighL := TRUE;                    // 高浓锁存
        _iFailCnt := _iFailCnt + 1;         // 连续失效计数加一
        _eState := E_DL_JbsCausticConcState.eJbsConcHigh;
    ELSIF _bLowRaw THEN
        _uInfo := 16#0091_0411;             // 信息级：接近下限但尚在去抖窗内
    ELSE
        _uInfo := 16#0091_0414;             // 信息级：浓度合格
        _iFailCnt := 0;                     // 回到带内即清连续失效计数
    END_IF

E_DL_JbsCausticConcState.eJbsConcLow:
    IF _iFailCnt >= fFailMax THEN
        _uFault := 16#0091_0415;            // 故障级：连续失效计数达上限（联动无效）
        _bLowL := FALSE;                    // 低浓锁存升格为故障，避免双码并存
        _bFault := TRUE;                    // 故障锁存
        _eState := E_DL_JbsCausticConcState.eJbsConcFault;
    ELSIF rtReset.Q THEN
        _bLowL := FALSE;                    // 解除路径：复位上升沿（可达，R188）
        _uFault := 16#0000_0000;            // 清锁存码
        _eState := E_DL_JbsCausticConcState.eJbsConcNormal;
    ELSIF NOT _bLowRaw AND NOT _bHighRaw THEN
        _bLowL := FALSE;                    // 浓度自行回到带内：清锁存（保留计数供累计判据）
        _eState := E_DL_JbsCausticConcState.eJbsConcNormal;
    END_IF

E_DL_JbsCausticConcState.eJbsConcHigh:
    IF _iFailCnt >= fFailMax THEN
        _uFault := 16#0091_0415;            // 故障级：连续失效计数达上限（联动无效）
        _bHighL := FALSE;                   // 高浓锁存升格为故障，避免双码并存
        _bFault := TRUE;                    // 故障锁存
        _eState := E_DL_JbsCausticConcState.eJbsConcFault;
    ELSIF rtReset.Q THEN
        _bHighL := FALSE;                   // 解除路径：复位上升沿（可达，R188）
        _uFault := 16#0000_0000;            // 清锁存码
        _eState := E_DL_JbsCausticConcState.eJbsConcNormal;
    ELSIF NOT _bLowRaw AND NOT _bHighRaw THEN
        _bHighL := FALSE;                   // 浓度自行回到带内：清锁存（保留计数供累计判据）
        _eState := E_DL_JbsCausticConcState.eJbsConcNormal;
    END_IF

E_DL_JbsCausticConcState.eJbsConcFault:
    IF rtReset.Q AND (NOT xFault) AND _bFinOk AND _bCfgOk THEN
        _bFault := FALSE;                   // 解除路径：复位沿 + 外部故障消失 + 入参/组态合法（可达，R188）
        _uFault := 16#0000_0000;            // 清锁存码
        _iFailCnt := 0;                     // 累计计数一并清（故障已人工确认）
        _eState := E_DL_JbsCausticConcState.eJbsConcNormal;
    END_IF

ELSE
    _uFault := 16#0091_0418;                // 故障级：非法相位 ID 兜底
    _bFault := TRUE;                        // 锁存
    _bLowL := FALSE;                        // 各级锁存清
    _bHighL := FALSE;
    _eState := E_DL_JbsCausticConcState.eJbsConcFault;        // 强制回故障相

END_CASE

(* —— 段 6：后置段（计数器域兜底：负值归零、越上限钳制，防整型溢出） —— *)
IF _iFailCnt < 0 THEN
    _iFailCnt := 0;                         // 负计数属异常，归零
END_IF
IF _iFailCnt > DL_CNT_HI THEN
    _iFailCnt := DL_CNT_HI;                 // 越上限钳制
END_IF

(* —— 段 7：出口单点映射（名实同源；请求位由状态导出，故障侧全清） —— *)
xLowAlarm := _bLowL AND (NOT _bFault);                                     // 低浓报警出口
xHighAlarm := _bHighL AND (NOT _bFault);                                   // 高浓报警出口
xMakeupReq := (_eState = E_DL_JbsCausticConcState.eJbsConcLow) AND (NOT _bFault);    // 补碱请求
xDiluteReq := (_eState = E_DL_JbsCausticConcState.eJbsConcHigh) AND (NOT _bFault);   // 稀释请求
nFailCount := _iFailCnt;                                                   // 计数出口
eState := _eState;                                                         // 状态出口单点映射
IF _bFault OR _bLowL OR _bHighL THEN
    nErrId := _uFault;                      // 故障码锁存回放（不在故障相按当下输入重推断）
ELSE
    nErrId := _uInfo;                       // 信息码
END_IF

END_FUNCTION_BLOCK

(* ---- FB_DL_ModuleLamVacuumSeq.st ---- *)
(*
  FB_DL_ModuleLamVacuumSeq  —  组件层压真空顺控（抽气-加热-加压-放气）/ Module laminator vacuum sequence
  分类 Category : DL_Process
  码位 Code     : 16#06_0_B5
  版本 Version  : 1.0.2
  来源 Source   : t2-7-packml — IEC 61131-3 标准语义的道莅防御性实现
  溯源 Origin   : clean-room 实现，层压工艺 PackML 段序公开语义借鉴，未复制任何源码行（RESUME 承接 R36 §4 #20 规格）
                  （段序语义对齐 FB_DL_StepSequencer，不实例化；三接口契约按 I_DL_* 真实成员名调用）
  功能 Function : 1) 四段顺控 Evac→Heat→Press→Vent，每段带 tSegmentTimeout 超时升级；
                  2) 加压段须真空度与温度双到位才允许升压（联锁内置，规格强制）；
                  3) 放气段结束须真空度回到常压确认（fVacKpa <= fAtmVacKpa）才进 Done；
                  4) 真空深度出口 fVacKpa = −iVac.fPressure（接口契约为负压值，出口取正深度）。
  边界 Boundary : ① 任一注入接口未装配校验由上层装配点承载（库内既有体例，__ISVALIDREF 为禁用项）；
                  ② 注入件 bFault（真空/温区/气缸）判故障升级；
                  ③ fPressTargetBar 超组态上限 fPressMaxBar 钳制并置信息码；配方四段全 0 判组态错；
                  ④ CASE 全态覆盖 + ELSE 兜底置 Fault；
                  ⑤ 解除式自证：bSegmentTimeoutFault 解除 = bReset 上升沿 AND eState = Idle；Idle 可达路径 =
                     每段正常推进（Evac→Heat→Press→Vent→Done→Idle）+ 超时 Fault 经 bReset 回 Idle，两条均给出；
                  ⑥ 段推进单发命令：各相进入拍单发一次（_bCmdLatch 承载，防重复下发）。
  依赖 Depends  : I_DL_VacuumGenerator / I_DL_TemperatureZone / I_DL_Cylinder（注入，不实例化）；
                  段序语义对齐 FB_DL_StepSequencer（已注册，不实例化）
  码表 Error codes（本件格 06_0_B5，子码步进 +0x100）:
    16#0006_01B5 信息级：周期完成（Done 相）
    16#0006_02B5 故障级：组态非法（目标 <= 0 / 配方全 0 / 超时 <= 0 / 上限 <= 0），锁存至复位
    16#0006_03B5 故障级：段超时升级（锁存，解除 = bReset 上升沿经 eFault 相迁出回 eIdle）
    16#0006_04B5 信息级：加压段真空联锁未满足（等待，不置故障）
    16#0006_05B5 故障级：注入件故障（真空/温区/气缸 bFault），锁存至复位
    16#0006_06B5 故障级：状态机落 ELSE 兜底（非法相位 ID）
    16#0006_07B5 信息级：压力目标越上限，已钳制

R39 返修（R38 终审挂账闭环，v1.0.2）: ① tonSeg PT 误接 tSegmentTimeout → 拆分为四相独立配方 TON
  （tonEvac/tonHeat/tonPress/tonVent，PT 各接本段配方时长，IN 单相等式，跨相迁移拍必断，R228-A 达标）；
  ② tonSegMax 跨相不复位 → 同步拆分为四相独立超时 TON（tonEvacTo/tonHeatTo/tonPressTo/tonVentTo）；
  ③ eFault 无迁出 → eFault 相新增 bReset 上升沿迁出边回 eIdle（迁出条件 = 输入引脚 rtReset.Q，恒可达）。
  修订历史 Revision :
    2026-11-19  v1.0.2  R39 返修：配方时长接入 + 相独立超时 + eFault 迁出边（R38 挂账三项闭环）
    2026-11-18  v1.0.0  R38 首版
*)

TYPE E_DL_LamPhase :
(
    eIdle  := 0,     // 空闲：等启动指令 / Idle, waiting for start
    eEvac  := 10,    // 抽气段 / Evacuation segment
    eHeat  := 20,    // 加热段 / Heating segment
    ePress := 30,    // 加压段（真空+温度双联锁）/ Pressing segment, dual interlock
    eVent  := 40,    // 放气段 / Venting segment
    eDone  := 50,    // 完成：常压确认落定 / Done, atmospheric confirmed
    eFault := 90     // 故障：组态/超时/注入件锁定 / Fault, latched
);
END_TYPE

FUNCTION_BLOCK FB_DL_ModuleLamVacuumSeq
VAR_INPUT
    bStart          : BOOL := FALSE;      // 启动指令（上升沿）/ Start command
    fVacTargetKpa   : REAL := 85.0;       // 真空目标深度 [kPa]，域 > 0 / Vacuum target depth
    fPressTargetBar : REAL := 1.5;        // 加压目标 [bar]，域 (0, fPressMaxBar] / Press target
    fPressMaxBar    : REAL := 2.0;        // 加压组态上限 [bar]，域 > 0 / Press ceiling
    fTempTargetC    : REAL := 145.0;      // 加热目标温度 [°C]，域 > 0 / Heating target temperature
    fAtmVacKpa      : REAL := 2.0;        // 常压确认阈值 [kPa]，域 >= 0 / Atmospheric confirmation threshold
    atEvacMs        : TIME := T#60S;      // 抽气段配方时长 [ms] / Evacuation recipe duration
    atHeatMs        : TIME := T#180S;     // 加热段配方时长 [ms] / Heating recipe duration
    atPressMs       : TIME := T#300S;     // 加压段配方时长 [ms] / Pressing recipe duration
    atVentMs        : TIME := T#30S;      // 放气段配方时长 [ms] / Venting recipe duration
    tSegmentTimeout : TIME := T#420S;     // 单段超时 [ms]，域 > 0 / Segment timeout
    bReset          : BOOL := FALSE;      // 复位（超时/故障解除路径之一）/ Reset
END_VAR
VAR_OUTPUT
    bCycleDone            : BOOL;         // 周期完成 / Cycle done
    bSegmentTimeoutFault  : BOOL;         // 段超时故障锁存（解除 = bReset AND Idle）/ Segment timeout latch
    nSegment              : INT;          // 当前段号 [0..3]（0=抽 1=热 2=压 3=放）/ Segment index
    fVacKpa               : REAL;         // 真空深度出口 [kPa]（取正深度）/ Vacuum depth outlet
    nErrId                : UDINT;        // 事件码，0 = 无事件 / Event code
    eState                : E_DL_LamPhase;// 状态出口，段尾单点映射 / State outlet
END_VAR
VAR_IN_OUT
    iVac      : I_DL_VacuumGenerator;     // 真空发生器引用（注入，不实例化）/ Vacuum reference
    iTempZone : I_DL_TemperatureZone;     // 温区引用（注入，不实例化）/ Temperature zone reference
    iPressCyl : I_DL_Cylinder;            // 压合气缸引用（注入，不实例化）/ Press cylinder reference
END_VAR
VAR
    tonEvac     : TON;                    // 抽气段配方计时（单相独占，PT=配方时长）/ Evacuation recipe timer
    tonHeat     : TON;                    // 加热段配方计时（单相独占，PT=配方时长）/ Heating recipe timer
    tonPress    : TON;                    // 加压段配方计时（单相独占，PT=配方时长）/ Pressing recipe timer
    tonVent     : TON;                    // 放气段配方计时（单相独占，PT=配方时长）/ Venting recipe timer
    tonEvacTo   : TON;                    // 抽气段超时（单相独占）/ Evacuation timeout
    tonHeatTo   : TON;                    // 加热段超时（单相独占）/ Heating timeout
    tonPressTo  : TON;                    // 加压段超时（单相独占）/ Pressing timeout
    tonVentTo   : TON;                    // 放气段超时（单相独占）/ Venting timeout
    tonFaultWch : TON;                    // 故障观察窗，自复位 / Fault watch window, self-resetting
    rtStart     : R_TRIG;                 // 启动上升沿 / Start rising edge
    rtReset     : R_TRIG;                 // 复位上升沿 / Reset rising edge
    _eState     : E_DL_LamPhase := E_DL_LamPhase.eIdle;   // 内部相位（CASE 唯一写入目标）/ Internal phase
    _bCmdLatch  : BOOL;                   // 本相命令已单发标志 / Phase command one-shot latch
    _rPressTgt  : REAL;                   // 钳制后压力目标 [bar] / Clamped press target
    _rTempAct   : REAL;                   // 温区实测温度 [°C] / Zone actual temperature
    _rVacDepth  : REAL;                   // 真空深度暂存 [kPa] / Vacuum depth scratch
    _bVacOk     : BOOL;                   // 真空到位标志 / Vacuum in-position flag
    _bTempOk    : BOOL;                   // 温度到位标志 / Temperature in-position flag
    _bToL       : BOOL;                   // 段超时锁存保持量 / Segment timeout latch
    _uFault     : UDINT;                  // 故障码锁存 / Latched fault code
    _uInfo      : UDINT;                  // 信息码，每拍重算 / Info code
    _bFault     : BOOL;                   // 故障锁存位 / Latched fault bit
    _bCfgBad    : BOOL;                   // 组态非法聚合 / Configuration invalid aggregate
END_VAR
VAR CONSTANT
    DL_SEG_EVAC  : INT := 0;    // 段号：抽气 / Segment index evacuation
    DL_SEG_HEAT  : INT := 1;    // 段号：加热 / Segment index heating
    DL_SEG_PRESS : INT := 2;    // 段号：加压 / Segment index pressing
    DL_SEG_VENT  : INT := 3;    // 段号：放气 / Segment index venting
    DL_WATCH_PT  : TIME := T#2S;   // 故障观察窗 [ms]，自复位 / Fault watch window
END_VAR

(* —— 段 0：定时器与边沿无条件周期刷新（R182：调用语句不得置于 IF/CASE 内） —— *)
rtStart(CLK := bStart);                                          // 启动上升沿，每拍必调
rtReset(CLK := bReset);                                          // 复位上升沿，每拍必调
tonFaultWch(IN := (NOT tonFaultWch.Q), PT := DL_WATCH_PT);       // 观察窗自复位（表达式入参）
tonEvac(IN := (_eState = E_DL_LamPhase.eEvac), PT := atEvacMs);      // 抽气配方计时（单相独占，PT=配方时长）
tonHeat(IN := (_eState = E_DL_LamPhase.eHeat), PT := atHeatMs);      // 加热配方计时（单相独占，PT=配方时长）
tonPress(IN := (_eState = E_DL_LamPhase.ePress), PT := atPressMs);   // 加压配方计时（单相独占，PT=配方时长）
tonVent(IN := (_eState = E_DL_LamPhase.eVent), PT := atVentMs);      // 放气配方计时（单相独占，PT=配方时长）
tonEvacTo(IN := (_eState = E_DL_LamPhase.eEvac), PT := tSegmentTimeout);    // 抽气段超时（单相独占）
tonHeatTo(IN := (_eState = E_DL_LamPhase.eHeat), PT := tSegmentTimeout);    // 加热段超时（单相独占）
tonPressTo(IN := (_eState = E_DL_LamPhase.ePress), PT := tSegmentTimeout);  // 加压段超时（单相独占）
tonVentTo(IN := (_eState = E_DL_LamPhase.eVent), PT := tSegmentTimeout);    // 放气段超时（单相独占）

(* —— 段 1：单拍量预清零（锁存量 _uFault/_bFault/_bToL/_bCmdLatch 不入清单，R187①） —— *)
_uInfo := 16#0000_0000;         // 信息码每拍重算
bCycleDone := FALSE;            // 完成出口缺省 FALSE（Done 相单点置位）
_bCfgBad := FALSE;              // 组态非法预清零
nErrId := 16#0000_0000;         // 事件码缺省无事件

(* —— 段 2：组态域闸（覆盖全部参与判据换算的引脚，R151） —— *)
IF (fVacTargetKpa <> fVacTargetKpa) OR (fVacTargetKpa <= 0.0)
   OR (fTempTargetC <> fTempTargetC) OR (fTempTargetC <= 0.0) THEN
    _bCfgBad := TRUE;           // 目标非法
END_IF
IF (fPressMaxBar <= 0.0) OR (fAtmVacKpa < 0.0) OR (TIME_TO_DINT(tSegmentTimeout) <= 0) THEN
    _bCfgBad := TRUE;           // 上限/常压阈/超时非法
END_IF
IF (TIME_TO_DINT(atEvacMs) <= 0) AND (TIME_TO_DINT(atHeatMs) <= 0)
   AND (TIME_TO_DINT(atPressMs) <= 0) AND (TIME_TO_DINT(atVentMs) <= 0) THEN
    _bCfgBad := TRUE;           // 配方四段全 0（规格强制）
END_IF

(* —— 段 3：复位沿（超时/故障解除式：bReset AND eState = Idle） —— *)
IF rtReset.Q THEN
    IF _eState = E_DL_LamPhase.eIdle THEN
        _bFault := FALSE;       // 清故障锁存位（Idle 可达，规格解除式）
        _uFault := 16#0000_0000;
        _bToL   := FALSE;       // 超时锁存清零
        bSegmentTimeoutFault := FALSE;
    END_IF
END_IF

(* —— 段 4：过程量只读采集与换算 —— *)
_rTempAct := iTempZone.fTempActual;          // 温区实测 [°C]
_rVacDepth := -iVac.fPressure;               // 真空深度 = 负压反馈取反 [kPa]（接口契约：负值=真空）
fVacKpa := _rVacDepth;                       // 深度出口（正深度）
_bVacOk := _rVacDepth >= fVacTargetKpa;      // 真空到位判据（每拍重算）
_bTempOk := ABS(_rTempAct - fTempTargetC) <= MAX(fTempTargetC * 0.02, 2.0);   // 温度到位（±2% 或 ±2°C 宽容）

(* —— 段 5：相位机（只做迁移与单发命令；出口在段 8） —— *)
CASE _eState OF

E_DL_LamPhase.eIdle:
    IF _bCfgBad THEN
        _uFault := 16#0006_02B5;            // 故障级：组态非法
        _bFault := TRUE;                    // 锁存（复位沿 + Idle 可清）
        _eState := E_DL_LamPhase.eFault;
    ELSIF rtStart.Q THEN
        IF fPressTargetBar > fPressMaxBar THEN
            _rPressTgt := fPressMaxBar;     // 压力目标越上限钳制
            _uInfo := 16#0006_07B5;         // 信息级：已钳制
        ELSE
            _rPressTgt := fPressTargetBar;  // 域内直通
        END_IF
        _bCmdLatch := FALSE;                // 命令单发标志复位
        iVac.CmdEvacuate();                 // 单发抽气指令
        iTempZone.CmdEnable(bOn := TRUE);   // 温区投运
        _bCmdLatch := TRUE;                 // 单发标志
        _eState := E_DL_LamPhase.eEvac;     // 进抽气段
    END_IF

E_DL_LamPhase.eEvac:
    IF (iVac.bFault OR iTempZone.bFault OR iPressCyl.bFault) THEN
        _uFault := 16#0006_05B5;            // 故障级：注入件故障
        _bFault := TRUE;
        iVac.CmdStop();                     // 安全侧全停
        iTempZone.CmdEnable(bOn := FALSE);
        _eState := E_DL_LamPhase.eFault;
    ELSIF tonEvacTo.Q THEN
        _bToL := TRUE;                      // 超时锁存
        _uFault := 16#0006_03B5;            // 故障级：段超时升级
        _bFault := TRUE;
        iVac.CmdStop();
        iTempZone.CmdEnable(bOn := FALSE);
        _eState := E_DL_LamPhase.eFault;
    ELSIF _bVacOk AND (TIME_TO_DINT(atEvacMs) <= 0 OR tonEvac.Q) THEN
        iTempZone.SetSetpoint(fTemp := fTempTargetC);   // 单发设定点
        _eState := E_DL_LamPhase.eHeat;     // 进加热段（正常推进，Idle 路径之一）
        _bCmdLatch := FALSE;
    END_IF

E_DL_LamPhase.eHeat:
    IF (iVac.bFault OR iTempZone.bFault OR iPressCyl.bFault) THEN
        _uFault := 16#0006_05B5;
        _bFault := TRUE;
        iVac.CmdStop();
        iTempZone.CmdEnable(bOn := FALSE);
        _eState := E_DL_LamPhase.eFault;
    ELSIF tonHeatTo.Q THEN
        _bToL := TRUE;
        _uFault := 16#0006_03B5;
        _bFault := TRUE;
        iVac.CmdStop();
        iTempZone.CmdEnable(bOn := FALSE);
        _eState := E_DL_LamPhase.eFault;
    ELSIF _bTempOk AND (TIME_TO_DINT(atHeatMs) <= 0 OR tonHeat.Q) THEN
        iPressCyl.CmdExtend();              // 单发升压
        _eState := E_DL_LamPhase.ePress;    // 进加压段
        _bCmdLatch := FALSE;
    END_IF

E_DL_LamPhase.ePress:
    IF (iVac.bFault OR iTempZone.bFault OR iPressCyl.bFault) THEN
        _uFault := 16#0006_05B5;
        _bFault := TRUE;
        iPressCyl.CmdStop();
        iVac.CmdStop();
        iTempZone.CmdEnable(bOn := FALSE);
        _eState := E_DL_LamPhase.eFault;
    ELSIF tonPressTo.Q THEN
        _bToL := TRUE;
        _uFault := 16#0006_03B5;
        _bFault := TRUE;
        iPressCyl.CmdStop();
        iVac.CmdStop();
        iTempZone.CmdEnable(bOn := FALSE);
        _eState := E_DL_LamPhase.eFault;
    ELSIF NOT (_bVacOk AND _bTempOk) THEN
        _uInfo := 16#0006_04B5;             // 信息级：真空/温度双联锁未满足（等待，不置故障）
    ELSIF iPressCyl.bExtended AND (TIME_TO_DINT(atPressMs) <= 0 OR tonPress.Q) THEN
        iVac.CmdBlowOff();                  // 单发放气
        _eState := E_DL_LamPhase.eVent;     // 进放气段
        _bCmdLatch := FALSE;
    END_IF

E_DL_LamPhase.eVent:
    IF (iVac.bFault OR iTempZone.bFault OR iPressCyl.bFault) THEN
        _uFault := 16#0006_05B5;
        _bFault := TRUE;
        iVac.CmdStop();
        iTempZone.CmdEnable(bOn := FALSE);
        _eState := E_DL_LamPhase.eFault;
    ELSIF tonVentTo.Q THEN
        _bToL := TRUE;
        _uFault := 16#0006_03B5;
        _bFault := TRUE;
        iVac.CmdStop();
        iTempZone.CmdEnable(bOn := FALSE);
        _eState := E_DL_LamPhase.eFault;
    ELSIF (_rVacDepth <= fAtmVacKpa) AND (TIME_TO_DINT(atVentMs) <= 0 OR tonVent.Q) THEN
        iTempZone.CmdEnable(bOn := FALSE);  // 温区退出
        iPressCyl.CmdRetract();             // 压头缩回
        _eState := E_DL_LamPhase.eDone;     // 常压确认：进完成相
    END_IF

E_DL_LamPhase.eDone:
    bCycleDone := TRUE;                     // 完成出口（Done 相每拍重申）
    _uInfo := 16#0006_01B5;                 // 信息级：周期完成
    IF NOT bStart THEN
        _eState := E_DL_LamPhase.eIdle;     // 指令撤销：回空闲（Idle 可达路径：正常推进链末端）
    END_IF

E_DL_LamPhase.eFault:
    IF rtReset.Q THEN                       // 迁出边：bReset 上升沿（R228-B：输入引脚，恒可达）
        _bFault := FALSE;                   // 清故障锁存位
        _uFault := 16#0000_0000;            // 清锁存码
        _bToL   := FALSE;                   // 超时锁存清零
        bSegmentTimeoutFault := FALSE;      // 超时出口同步清除
        _eState := E_DL_LamPhase.eIdle;     // 迁出：回空闲（Idle 可达路径：故障迁出边）
    END_IF

ELSE
    _uFault := 16#0006_06B5;                // 故障级：非法相位 ID 兜底
    _bFault := TRUE;                        // 锁存
    _eState := E_DL_LamPhase.eFault;        // 强制回故障相

END_CASE

(* —— 段 6：出口单点映射（名实同源；锁存码回放，禁同拍抹除） —— *)
IF _eState = E_DL_LamPhase.eEvac THEN
    nSegment := DL_SEG_EVAC;                // 段号 0：抽气
ELSIF _eState = E_DL_LamPhase.eHeat THEN
    nSegment := DL_SEG_HEAT;                // 段号 1：加热
ELSIF _eState = E_DL_LamPhase.ePress THEN
    nSegment := DL_SEG_PRESS;               // 段号 2：加压
ELSIF _eState = E_DL_LamPhase.eVent THEN
    nSegment := DL_SEG_VENT;                // 段号 3：放气
ELSE
    nSegment := -1;                         // Idle/Done/Fault：无有效段号
END_IF
bSegmentTimeoutFault := _bToL;              // 超时出口 = 锁存量（置位同拍不被抹）
IF _bFault THEN
    nErrId := _uFault;          // 故障锁存码回放（不在故障相按当下输入重推）
    bCycleDone := FALSE;        // 故障相完成出口强制 FALSE（安全侧）
ELSE
    nErrId := _uInfo;           // 信息码
END_IF
eState := _eState;              // 状态出口单点映射

END_FUNCTION_BLOCK
